// TwinCAT 3 PLC project TwinCAT_OpenFramework_Testing
// Title: TwinCAT Open Framework Testing
// Company: Oleksandr Tiutyk FOP
// Author: Oleksandr Tiutyk
// ProjectVersion: 1.0.13.0
// Description: Auumated testing engine implemenation
// ProgramVersion: 3.1.4026.28
// libraries:
//   Tc2_Utilities, * (Beckhoff Automation GmbH)
//   [TwinCAT Open Framework Core], * (Oleksandr Tiutyk FOP)
// project tree:
//   Assertions/ Assertions.TcPOU, AssertionContext.TcPOU
//   Assertions/TypedContexts/ BoolAssertionContext.TcPOU, SIntAssertionContext.TcPOU, IntAssertionContext.TcPOU, DIntAssertionContext.TcPOU, LIntAssertionContext.TcPOU, USIntAssertionContext.TcPOU, UIntAssertionContext.TcPOU, UDIntAssertionContext.TcPOU, ULIntAssertionContext.TcPOU, ByteAssertionContext.TcPOU, WordAssertionContext.TcPOU, DWordAssertionContext.TcPOU, LWordAssertionContext.TcPOU, RealAssertionContext.TcPOU, LongRealAssertionContext.TcPOU, StringAssertionContext.TcPOU, WideStringAssertionContext.TcPOU, TimeAssertionContext.TcPOU, LongTimeAssertionContext.TcPOU, DateAssertionContext.TcPOU, LongDateAssertionContext.TcPOU, DateTimeAssertionContext.TcPOU, LongDateTimeAssertionContext.TcPOU, TimeOfDayAssertionContext.TcPOU, LongTimeOfDayAssertionContext.TcPOU, PointerAssertionContext.TcPOU
//   Internal/ CurrentNamespace.TcPOU, NamespaceExtractor.TcPOU
//   Runner/ TEST_RUN_PHASE.TcDUT, TestRunner.TcPOU
//   TestElements/Groups/ TestGroup.TcPOU
//   TestElements/ IParentTestElement.TcIO, TEST_ELEMENT_STATE.TcDUT, ITestElement.TcIO, TestElement.TcPOU
//   TestElements/Tests/ TEST_CYCLE_RESULT.TcDUT, TEST_OUTCOME.TcDUT, ITestCase.TcIO, TestCase.TcPOU, SingleCycleTest.TcPOU, MultiCycleTest.TcPOU
//   Reporting/ ITestReporter.TcIO, AdsLogReporter.TcPOU, JUnitXmlReporter.TcPOU
//   / TestServices.TcPOU
//   Version/ Global_Version.TcGVL
// (motion and I/O tree: see PLC project twincat_openframework_core)
// real-time tasks:
//   TASK PlcTask: cycle T#10ms, priority 20, ADS port 350
//   TASK TestTask: cycle T#10ms, priority 1, ADS port 351
//   TASK RunnerTestTask: cycle T#10ms, priority 2, ADS port 354
//   TASK HowToTask: cycle T#10ms, priority 22, ADS port 353
// variable links:

// ---- Runner/TEST_RUN_PHASE.TcDUT
(*
SPDX-FileCopyrightText: © 2026 Oleksandr Tiutyk <trofimich@gmail.com>
SPDX-License-Identifier: MIT
License: https://opensource.org/license/mit
*)

(*!
<summary>Identifies the next root scheduling or reporting action.</summary>
*)

{attribute 'qualified_only'}
{attribute 'strict'}
{attribute 'to_string'}
TYPE TEST_RUN_PHASE :
(
	STARTING,
	RUNNING_ELEMENTS,
	REPORTING_TOTALS,
	COMPLETED
);
END_TYPE

// ---- TestElements/Tests/TEST_CYCLE_RESULT.TcDUT
(*
SPDX-FileCopyrightText: © 2026 Oleksandr Tiutyk <trofimich@gmail.com>
SPDX-License-Identifier: MIT
License: https://opensource.org/license/mit
*)

(*!
<summary>Indicates whether a test body needs more scheduling cycles or has finished on the current cycle.</summary>
<description>
BUSY (0) is the default uninitialized value and keeps the test running across subsequent cycles unless a failure
or deadline terminates the run. DONE (1) requests normal completion after the current cycle returns.
</description>
*)

{attribute 'qualified_only'}
{attribute 'strict'}
{attribute 'to_string'}
TYPE TEST_CYCLE_RESULT :
(
	BUSY := 0,
	DONE := 1
);
END_TYPE

// ---- TestElements/Tests/TEST_OUTCOME.TcDUT
(*
SPDX-FileCopyrightText: © 2026 Oleksandr Tiutyk <trofimich@gmail.com>
SPDX-License-Identifier: MIT
License: https://opensource.org/license/mit
*)

(*!
<summary>Defines the execution outcome of an individual test scenario.</summary>
<description>
Tracks whether a test has not yet run, is currently executing across cycles, passed all assertions, failed an
assertion or invariant, or was explicitly skipped.
</description>
*)

{attribute 'qualified_only'}
{attribute 'strict'}
{attribute 'to_string'}
TYPE TEST_OUTCOME :
(
	NOT_RUN := 0,
	RUNNING := 1,
	PASSED := 2,
	FAILED := 3,
	SKIPPED := 4
);
END_TYPE

// ---- TestElements/TEST_ELEMENT_STATE.TcDUT
(*
SPDX-FileCopyrightText: © 2026 Oleksandr Tiutyk <trofimich@gmail.com>
SPDX-License-Identifier: MIT
License: https://opensource.org/license/mit
*)

(*!
<summary>Identifies the execution lifecycle of a test element.</summary>
*)

{attribute 'qualified_only'}
{attribute 'strict'}
{attribute 'to_string'}
TYPE TEST_ELEMENT_STATE :
(
	READY,
	RUNNING,
	COMPLETED
);
END_TYPE

// ---- Version/Global_Version.TcGVL
{attribute 'TcGenerated'}
{attribute 'no-analysis'}
{attribute 'linkalways'}
// This function has been automatically generated from the project information.
VAR_GLOBAL CONSTANT
	{attribute 'const_non_replaced'}
	stLibVersion_TwinCAT_Open_Framework_Testing : ST_LibVersion := (iMajor := 1, iMinor := 0, iBuild := 13, iRevision := 0, nFlags := 0, sVersion := '1.0.13.0');
END_VAR

// ---- TestElements/IParentTestElement.TcIO
(*
SPDX-FileCopyrightText: © 2026 Oleksandr Tiutyk <trofimich@gmail.com>
SPDX-License-Identifier: MIT
License: https://opensource.org/license/mit
*)

(*!
<summary>Exposes borrowed direct children of a test element in fixed execution order.</summary>
<description>
ChildCount is stable throughout the element's lifetime; each direct child occupies one non-null slot.
GetChildByIndex borrows a child without resetting or executing it and transfers no allocation ownership.
Children and parent links obey ITestElement lifetime and lifecycle rules. Observations belong to the owning
task without reentry or cross-task synchronization. An empty composition has ChildCount zero and no valid index.
</description>
*)

INTERFACE IParentTestElement EXTENDS ITestElement

(*!
<summary>Reports the fixed number of direct children, including zero for an empty composition.</summary>
*)

{attribute 'monitoring' := 'call'}
PROPERTY FINAL ChildCount : TOF_Core.INT_LENGTH
GET
END_GET
END_PROPERTY

(*!
<summary>Borrows a direct child by its zero-based position in fixed execution order.</summary>
<description>
Available before the first Reset and after a failed Reset, provided the backing array and selected slot exist.
Missing storage or a null selected slot raises DataMemberNotSpecifiedException. Storage is checked first;
an index outside zero through ChildCount minus one raises ArgumentOutOfRangeException.
Does not mutate or execute the child, repeat whole-tree validation, or transfer ownership.
The child must remain alive while the interface is used; use only from the tree's owning task without reentry.
</description>
<param name="index">Zero-based direct-child position; an empty composition has no valid value.</param>
*)
METHOD GetChildByIndex : ITestElement
VAR_INPUT
	index : TOF_Core.INT_LENGTH;
END_VAR
END_METHOD

END_INTERFACE

// ---- Reporting/ITestReporter.TcIO
(*
SPDX-FileCopyrightText: © 2026 Oleksandr Tiutyk <trofimich@gmail.com>
SPDX-License-Identifier: MIT
License: https://opensource.org/license/mit
*)

(*!
<summary>Receives run boundaries and one terminal result per leaf test.</summary>
<description>
Callbacks execute synchronously in the owning runner task. Inputs are borrowed for the call only.
Do not retain them, reenter the tree, or share mutable reporter state between tasks. An exception aborts the
runner with ExitCode -1; output may be incomplete and the callback is not retried. Group paths are bounded
slash-separated display names. Groups do not emit synthetic test results or nested suite callbacks.
ReportTestCaseResult requires PASSED, FAILED or SKIPPED; other outcomes are invalid configuration.
Individual test names are bounded to 80 wide characters, matching INamed; group paths retain their 255-character bound.
</description>
*)

INTERFACE ITestReporter EXTENDS TOF_Core.IObject

(*!
<summary>Completes a run with aggregated leaf counts and nominal duration.</summary>
*)
METHOD ReportRunEnd
VAR_INPUT
	totalTests : TOF_Core.DINT_LENGTH;
	passedTests : TOF_Core.DINT_LENGTH;
	failedTests : TOF_Core.DINT_LENGTH;
	skippedTests : TOF_Core.DINT_LENGTH;
	duration : TIME;
END_VAR
END_METHOD

(*!
<summary>Begins a run with the number of configured leaf tests, including those that may be skipped.</summary>
<param name="testCount">The sum of the root TestCount values before executing any test.</param>
*)
METHOD ReportRunStart
VAR_INPUT
	testCount : TOF_Core.DINT_LENGTH;
END_VAR
END_METHOD

(*!
<summary>Receives one terminal leaf outcome and its first copied diagnostic.</summary>
<param name="testName">Individual name of at most 80 wide characters; longer input uses IEC truncation.</param>
*)
METHOD ReportTestCaseResult
VAR_INPUT
	groupPath : WSTRING(255);
	testName : WSTRING;
	outcome : TEST_OUTCOME;
	duration : TIME;
END_VAR
VAR_IN_OUT CONSTANT
	message : TOF_Core.ERROR_MESSAGE;
END_VAR
END_METHOD

END_INTERFACE

// ---- TestElements/ITestElement.TcIO
(*
SPDX-FileCopyrightText: © 2026 Oleksandr Tiutyk <trofimich@gmail.com>
SPDX-License-Identifier: MIT
License: https://opensource.org/license/mit
*)

(*!
<summary>Common cyclic execution contract for an individual test or a group of tests.</summary>
<description>
A live element occupies one slot of one tree. Its parent is assigned at construction and remains unchanged.
Its parent, descendants, reporter and tested resources remain alive and stable during a run.
All execution, configuration and observation of a tree belong to one cyclic task without reentry.
Separate tasks use disjoint trees, reporters and mutable tested resources; this interface provides no synchronization.
Execute advances at most one leaf body per call. A completed element ignores Execute until Reset.
Outcome counters describe leaf results. TestCount describes the configured leaf population of the subtree.
Custom implementations must preserve parent links and all lifecycle rules; callback exceptions abort the runner.
</description>
*)

INTERFACE ITestElement EXTENDS TOF_Core.INamed, TOF_Core.IExecutable

(*!
<summary>Reports nominal execution duration accumulated from calling task periods.</summary>
*)
{attribute 'monitoring' := 'call'}
PROPERTY Duration : TIME
GET
END_GET
END_PROPERTY

(*!
<summary>Counts failed leaf tests in this element.</summary>
*)
{attribute 'monitoring' := 'call'}
PROPERTY FailedCount : TOF_Core.DINT_LENGTH
GET
END_GET
END_PROPERTY

(*!
<summary>Builds the full display path from the root through this element.</summary>
<description>
Joins nonempty names with '/', including this element's name. A nameless root returns an empty path.
The result is a copied WSTRING bounded to 255 characters; overflow preserves the root prefix and ends with an ellipsis.
Reads the live Parent and Name properties without caching or changing the tree. All providers must remain alive
and stable during the call; use only in the owning task without reentry. Can be called before Reset.
A cyclic Parent chain raises StandardException to prevent an endless traversal. Provider exceptions propagate;
no element state or ownership is changed. Valid traversal uses fixed local strings without recursion or heap allocation.
</description>
*)
METHOD GetPath : WSTRING(255)
END_METHOD

(*!
<summary>Reports whether this element has completed.</summary>
*)
{attribute 'monitoring' := 'call'}
PROPERTY IsFinished : BOOL
GET
END_GET
END_PROPERTY

(*!
<summary>Reports whether this element has started and has not completed.</summary>
*)
{attribute 'monitoring' := 'call'}
PROPERTY IsRunning : BOOL
GET
END_GET
END_PROPERTY

(*!
<summary>Returns the group assigned at construction, or zero for a root.</summary>
<description>
Borrowed lifetime association. Reset and execution do not change it; the parent must remain alive.
Root registration with a runner does not bind Parent; a root must belong to one runner only.
</description>
*)
{attribute 'monitoring' := 'call'}
PROPERTY Parent : ITestElement
GET
END_GET
END_PROPERTY

(*!
<summary>Counts passed leaf tests in this element.</summary>
*)
{attribute 'monitoring' := 'call'}
PROPERTY PassedCount : TOF_Core.DINT_LENGTH
GET
END_GET
END_PROPERTY

(*!
<summary>Reports nominal scheduled duration, not CPU execution time.</summary>
*)
{attribute 'monitoring' := 'call'}
PROPERTY FINAL Reporter : ITestReporter
GET
END_GET
END_PROPERTY

(*!
<summary>Prepares a fresh run and borrows the reporter.</summary>
<description>
Call before first execution, after completion, or after an aborted run once resources are safe.
This is not cancellation: it does not execute test teardown. The reporter may be zero to suppress reporting.
Group reset recursively resets descendants. External callback exceptions propagate; partial reset is possible.
</description>
*)
METHOD Reset
VAR_INPUT
	reporter : ITestReporter;
END_VAR
END_METHOD

(*!
<summary>Counts skipped leaf tests in this element.</summary>
*)
{attribute 'monitoring' := 'call'}
PROPERTY SkippedCount : TOF_Core.DINT_LENGTH
GET
END_GET
END_PROPERTY

(*!
<summary>Reports nominal scheduled duration, not CPU execution time.</summary>
*)
{attribute 'monitoring' := 'call'}
PROPERTY FINAL State : TEST_ELEMENT_STATE
GET
END_GET
END_PROPERTY

(*!
<summary>Counts the configured leaf tests in this subtree.</summary>
<description>
A leaf counts as one regardless of its outcome. Groups sum their children; an empty group counts as zero.
Read from the owning task after the tree has been constructed. The caller supplies a valid, stable subtree
whose total fits in UDINT. Reading does not run or reset tests, and the value is stable across runs.
Provider exceptions propagate.
</description>
*)
{attribute 'monitoring' := 'call'}
PROPERTY TestCount : TOF_Core.DINT_LENGTH
GET
END_GET
END_PROPERTY

END_INTERFACE

// ---- TestElements/Tests/ITestCase.TcIO
(*
SPDX-FileCopyrightText: © 2026 Oleksandr Tiutyk <trofimich@gmail.com>
SPDX-License-Identifier: MIT
License: https://opensource.org/license/mit
*)

(*!
<summary>Receives assertion failures for one individual test.</summary>
<description>
Groups use ITestElement and do not receive leaf assertions. A failure is copied only while the case is running.
</description>
*)

INTERFACE ITestCase EXTENDS ITestElement

(*!
<summary>Copies the first failure of the running case; later diagnostics do not replace it.</summary>
*)
METHOD RecordFailure
VAR_IN_OUT CONSTANT
	message : TOF_Core.ERROR_MESSAGE;
END_VAR
END_METHOD

END_INTERFACE

// ---- Assertions/Assertions.TcPOU
(*
SPDX-FileCopyrightText: © 2026 Oleksandr Tiutyk <trofimich@gmail.com>
SPDX-License-Identifier: MIT
License: https://opensource.org/license/mit
*)

(*!
<summary>Provides fluent test assertion entry points on values, variables, and objects.</summary>
<description>
TestCase owns and binds this instance before its first callback.
Typed That methods copy actual values into independent persistent contexts; generic That borrows a live variable.
Contexts do not call one another; shared services only report failures and implement floating value policy.
Finish one immediate chain before starting another, regardless of operand type. Do not retain a returned
context or use this provider across tasks or reentrantly. Every entry verifies that its owning case is running.
An optional copied message prefixes every assertion failure in the chain and is replaced on the next entry.
Typed contexts apply ordinary IEC input conversions; select the entry matching the intended operand type.
Do not copy this provider by value: its contexts retain borrowed links to the owning test case and actual storage.
</description>
*)

{attribute 'no_explicit_call' := 'do not call this function block directly'}
FUNCTION_BLOCK Assertions EXTENDS TOF_Core.Object
VAR_STAT
	{attribute 'hide'} 
	_ClassName : STRING := __POUNAME();	
END_VAR
VAR	
	_AssertionContext : AssertionContext;
	
	_BoolContext : BoolAssertionContext;
	_SIntContext : SIntAssertionContext;
	_IntContext : IntAssertionContext;
	_DIntContext : DIntAssertionContext;
	_LIntContext : LIntAssertionContext;
	_USIntContext : USIntAssertionContext;
	_UIntContext : UIntAssertionContext;
	_UDIntContext : UDIntAssertionContext;
	_ULIntContext : ULIntAssertionContext;
	_ByteContext : ByteAssertionContext;
	_WordContext : WordAssertionContext;
	_DWordContext : DWordAssertionContext;
	_LWordContext : LWordAssertionContext;
	_RealContext : RealAssertionContext;
	_LongRealContext : LongRealAssertionContext;
	_StringContext : StringAssertionContext;
	_WideStringContext : WideStringAssertionContext;
	_TimeContext : TimeAssertionContext;
	_LongTimeContext : LongTimeAssertionContext;
	_DateContext : DateAssertionContext;
	_LongDateContext : LongDateAssertionContext;
	_DateTimeContext : DateTimeAssertionContext;
	_LongDateTimeContext : LongDateTimeAssertionContext;
	_TimeOfDayContext : TimeOfDayAssertionContext;
	_LongTimeOfDayContext : LongTimeOfDayAssertionContext;
	_PointerContext : PointerAssertionContext;
	
	_TestCase : ITestCase;
END_VAR

//! <summary>Borrows the owning test case for assertion failure reporting throughout the run.</summary>
METHOD INTERNAL FINAL Bind
VAR_INPUT
	testCase : ITestCase;
END_VAR
_TestCase := testCase;
END_METHOD

//! <summary>Provides assertion-provider metadata.</summary>
{attribute 'monitoring' := 'call'}
PROPERTY ClassName : REFERENCE TO STRING
GET
ClassName REF= _ClassName;
END_GET
END_PROPERTY

(*!
<summary>Returns the namespace name of this assertion provider.</summary>
*)
{attribute 'monitoring' := 'call'}
PROPERTY NamespaceName : REFERENCE TO STRING
GET
NamespaceName REF= CurrentNamespace.Name;
END_GET
END_PROPERTY

(*!
<summary>Rejects assertion entry outside a running owning case before context mutation.</summary>
<description>
Raises DataMemberNotSpecifiedException when no running test case is bound.
</description>
*)
METHOD PRIVATE requireRunningCase
IF _TestCase = 0 OR_ELSE NOT _TestCase.IsRunning THEN
	TOF_Core.Exceptions.ThrowDataMemberNotSpecified(
		sourceNamespaceName := NamespaceName,
		sourceClassName := ClassName,
		sourcePOUName := __POUNAME(),
		sourcePosition := __POSITION(),
		dataMemberName := '_TestCase'
	);
END_IF
END_METHOD

(*!
<summary>Reports the byte size of this concrete instance.</summary>
<description>
Uses XSIZEOF on the instance. Does not include separately allocated payloads or prove that an arbitrary
address is valid.
</description>
*)
{attribute 'monitoring' := 'call'}
PROPERTY SelfSize : ULINT
GET
SelfSize := XSIZEOF(THIS^);
END_GET
END_PROPERTY

(*!
<summary>Begins a fluent assertion chain on the provided actual value.</summary>
<description>
Borrows actual storage for this expression; actual must be a variable. Use typed entry points for literals
and expression results. Starting another chain replaces that entry's operand and message.
Calling That without a running owning case raises DataMemberNotSpecifiedException.
Equality follows GENERIC_VALUE byte/value semantics; FB operands do not invoke Object.Equals.
For object equality, use ThatBool on the Boolean result of its explicit Equals call.
</description>
<param name="actual">Live variable borrowed through the immediate chain.</param>
<param name="message">Optional copied prefix for every failure in this chain; default empty.</param>
*)
METHOD That : REFERENCE TO AssertionContext
VAR_INPUT
	actual : ANY;
	message : WSTRING(255) := "";
END_VAR
requireRunningCase();

_AssertionContext.Prepare(actual := actual, testCase := _TestCase, message := message);

That REF= _AssertionContext;
END_METHOD

(*!
<summary>Begins a fluent chain on a copied BOOL value.</summary>
<description>
Accepts literals, variables and expression results through a concrete IEC input type.
Requires a running owning case; otherwise raises DataMemberNotSpecifiedException.
Finish this chain before starting another. The message applies to every assertion in the chain.
</description>
<param name="actual">Value copied after ordinary IEC conversion to BOOL.</param>
<param name="message">Optional copied diagnostic prefix; default empty replaces the previous prefix.</param>
*)
METHOD ThatBool : REFERENCE TO BoolAssertionContext
VAR_INPUT
	actual : BOOL;
	message : WSTRING(255) := "";
END_VAR
requireRunningCase();

_BoolContext.Prepare(actual := actual, testCase := _TestCase, message := message);

ThatBool REF= _BoolContext;
END_METHOD

(*!
<summary>Begins a fluent chain on a copied BYTE value.</summary>
<description>
Accepts literals, variables and expression results through a concrete IEC input type.
Requires a running owning case; otherwise raises DataMemberNotSpecifiedException.
Finish this chain before starting another. The message applies to every assertion in the chain.
</description>
<param name="actual">Value copied after ordinary IEC conversion to BYTE.</param>
<param name="message">Optional copied diagnostic prefix; default empty replaces the previous prefix.</param>
*)
METHOD ThatByte : REFERENCE TO ByteAssertionContext
VAR_INPUT
	actual : BYTE;
	message : WSTRING(255) := "";
END_VAR
requireRunningCase();

_ByteContext.Prepare(actual := actual, testCase := _TestCase, message := message);

ThatByte REF= _ByteContext;
END_METHOD

(*!
<summary>Begins a fluent chain on a copied DATE value.</summary>
<description>
Accepts literals, variables and expression results through a concrete IEC input type.
Requires a running owning case; otherwise raises DataMemberNotSpecifiedException.
Finish this chain before starting another. The message applies to every assertion in the chain.
</description>
<param name="actual">Value copied after ordinary IEC conversion to DATE.</param>
<param name="message">Optional copied diagnostic prefix; default empty replaces the previous prefix.</param>
*)
METHOD ThatDate : REFERENCE TO DateAssertionContext
VAR_INPUT
	actual : DATE;
	message : WSTRING(255) := "";
END_VAR
requireRunningCase();

_DateContext.Prepare(actual := actual, testCase := _TestCase, message := message);

ThatDate REF= _DateContext;
END_METHOD

(*!
<summary>Begins a fluent chain on a copied DATE_AND_TIME value.</summary>
<description>
Accepts literals, variables and expression results through a concrete IEC input type.
Requires a running owning case; otherwise raises DataMemberNotSpecifiedException.
Finish this chain before starting another. The message applies to every assertion in the chain.
</description>
<param name="actual">Value copied after ordinary IEC conversion to DATE_AND_TIME.</param>
<param name="message">Optional copied diagnostic prefix; default empty replaces the previous prefix.</param>
*)
METHOD ThatDateTime : REFERENCE TO DateTimeAssertionContext
VAR_INPUT
	actual : DATE_AND_TIME;
	message : WSTRING(255) := "";
END_VAR
requireRunningCase();

_DateTimeContext.Prepare(actual := actual, testCase := _TestCase, message := message);

ThatDateTime REF= _DateTimeContext;
END_METHOD

(*!
<summary>Begins a fluent chain on a copied DINT value.</summary>
<description>
Accepts literals, variables and expression results through a concrete IEC input type.
Requires a running owning case; otherwise raises DataMemberNotSpecifiedException.
Finish this chain before starting another. The message applies to every assertion in the chain.
</description>
<param name="actual">Value copied after ordinary IEC conversion to DINT.</param>
<param name="message">Optional copied diagnostic prefix; default empty replaces the previous prefix.</param>
*)
METHOD ThatDInt : REFERENCE TO DIntAssertionContext
VAR_INPUT
	actual : DINT;
	message : WSTRING(255) := "";
END_VAR
requireRunningCase();

_DIntContext.Prepare(actual := actual, testCase := _TestCase, message := message);

ThatDInt REF= _DIntContext;
END_METHOD

(*!
<summary>Begins a fluent chain on a copied DWORD value.</summary>
<description>
Accepts literals, variables and expression results through a concrete IEC input type.
Requires a running owning case; otherwise raises DataMemberNotSpecifiedException.
Finish this chain before starting another. The message applies to every assertion in the chain.
</description>
<param name="actual">Value copied after ordinary IEC conversion to DWORD.</param>
<param name="message">Optional copied diagnostic prefix; default empty replaces the previous prefix.</param>
*)
METHOD ThatDWord : REFERENCE TO DWordAssertionContext
VAR_INPUT
	actual : DWORD;
	message : WSTRING(255) := "";
END_VAR
requireRunningCase();

_DWordContext.Prepare(actual := actual, testCase := _TestCase, message := message);

ThatDWord REF= _DWordContext;
END_METHOD

(*!
<summary>Begins a fluent chain on a copied INT value.</summary>
<description>
Accepts literals, variables and expression results through a concrete IEC input type.
Requires a running owning case; otherwise raises DataMemberNotSpecifiedException.
Finish this chain before starting another. The message applies to every assertion in the chain.
</description>
<param name="actual">Value copied after ordinary IEC conversion to INT.</param>
<param name="message">Optional copied diagnostic prefix; default empty replaces the previous prefix.</param>
*)
METHOD ThatInt : REFERENCE TO IntAssertionContext
VAR_INPUT
	actual : INT;
	message : WSTRING(255) := "";
END_VAR
requireRunningCase();

_IntContext.Prepare(actual := actual, testCase := _TestCase, message := message);

ThatInt REF= _IntContext;
END_METHOD

(*!
<summary>Begins a fluent chain on a copied LINT value.</summary>
<description>
Accepts literals, variables and expression results through a concrete IEC input type.
Requires a running owning case; otherwise raises DataMemberNotSpecifiedException.
Finish this chain before starting another. The message applies to every assertion in the chain.
</description>
<param name="actual">Value copied after ordinary IEC conversion to LINT.</param>
<param name="message">Optional copied diagnostic prefix; default empty replaces the previous prefix.</param>
*)
METHOD ThatLInt : REFERENCE TO LIntAssertionContext
VAR_INPUT
	actual : LINT;
	message : WSTRING(255) := "";
END_VAR
requireRunningCase();

_LIntContext.Prepare(actual := actual, testCase := _TestCase, message := message);

ThatLInt REF= _LIntContext;
END_METHOD

(*!
<summary>Begins a fluent chain on a copied LDATE value.</summary>
<description>
Accepts literals, variables and expression results through a concrete IEC input type.
Requires a running owning case; otherwise raises DataMemberNotSpecifiedException.
Finish this chain before starting another. The message applies to every assertion in the chain.
</description>
<param name="actual">Value copied after ordinary IEC conversion to LDATE.</param>
<param name="message">Optional copied diagnostic prefix; default empty replaces the previous prefix.</param>
*)
METHOD ThatLongDate : REFERENCE TO LongDateAssertionContext
VAR_INPUT
	actual : LDATE;
	message : WSTRING(255) := "";
END_VAR
requireRunningCase();

_LongDateContext.Prepare(actual := actual, testCase := _TestCase, message := message);

ThatLongDate REF= _LongDateContext;
END_METHOD

(*!
<summary>Begins a fluent chain on a copied LDATE_AND_TIME value.</summary>
<description>
Accepts literals, variables and expression results through a concrete IEC input type.
Requires a running owning case; otherwise raises DataMemberNotSpecifiedException.
Finish this chain before starting another. The message applies to every assertion in the chain.
</description>
<param name="actual">Value copied after ordinary IEC conversion to LDATE_AND_TIME.</param>
<param name="message">Optional copied diagnostic prefix; default empty replaces the previous prefix.</param>
*)
METHOD ThatLongDateTime : REFERENCE TO LongDateTimeAssertionContext
VAR_INPUT
	actual : LDATE_AND_TIME;
	message : WSTRING(255) := "";
END_VAR
requireRunningCase();

_LongDateTimeContext.Prepare(actual := actual, testCase := _TestCase, message := message);

ThatLongDateTime REF= _LongDateTimeContext;
END_METHOD

(*!
<summary>Begins a fluent chain on a copied LREAL value.</summary>
<description>
Accepts literals, variables and expression results through a concrete IEC input type.
Requires a running owning case; otherwise raises DataMemberNotSpecifiedException.
Finish this chain before starting another. The message applies to every assertion in the chain.
</description>
<param name="actual">Value copied after ordinary IEC conversion to LREAL.</param>
<param name="message">Optional copied diagnostic prefix; default empty replaces the previous prefix.</param>
*)
METHOD ThatLongReal : REFERENCE TO LongRealAssertionContext
VAR_INPUT
	actual : LREAL;
	message : WSTRING(255) := "";
END_VAR
requireRunningCase();

_LongRealContext.Prepare(actual := actual, testCase := _TestCase, message := message);

ThatLongReal REF= _LongRealContext;
END_METHOD

(*!
<summary>Begins a fluent chain on a copied LTIME value.</summary>
<description>
Accepts literals, variables and expression results through a concrete IEC input type.
Requires a running owning case; otherwise raises DataMemberNotSpecifiedException.
Finish this chain before starting another. The message applies to every assertion in the chain.
</description>
<param name="actual">Value copied after ordinary IEC conversion to LTIME.</param>
<param name="message">Optional copied diagnostic prefix; default empty replaces the previous prefix.</param>
*)
METHOD ThatLongTime : REFERENCE TO LongTimeAssertionContext
VAR_INPUT
	actual : LTIME;
	message : WSTRING(255) := "";
END_VAR
requireRunningCase();

_LongTimeContext.Prepare(actual := actual, testCase := _TestCase, message := message);

ThatLongTime REF= _LongTimeContext;
END_METHOD

(*!
<summary>Begins a fluent chain on a copied LTIME_OF_DAY value.</summary>
<description>
Accepts literals, variables and expression results through a concrete IEC input type.
Requires a running owning case; otherwise raises DataMemberNotSpecifiedException.
Finish this chain before starting another. The message applies to every assertion in the chain.
</description>
<param name="actual">Value copied after ordinary IEC conversion to LTIME_OF_DAY.</param>
<param name="message">Optional copied diagnostic prefix; default empty replaces the previous prefix.</param>
*)
METHOD ThatLongTimeOfDay : REFERENCE TO LongTimeOfDayAssertionContext
VAR_INPUT
	actual : LTIME_OF_DAY;
	message : WSTRING(255) := "";
END_VAR
requireRunningCase();

_LongTimeOfDayContext.Prepare(actual := actual, testCase := _TestCase, message := message);

ThatLongTimeOfDay REF= _LongTimeOfDayContext;
END_METHOD

(*!
<summary>Begins a fluent chain on a copied LWORD value.</summary>
<description>
Accepts literals, variables and expression results through a concrete IEC input type.
Requires a running owning case; otherwise raises DataMemberNotSpecifiedException.
Finish this chain before starting another. The message applies to every assertion in the chain.
</description>
<param name="actual">Value copied after ordinary IEC conversion to LWORD.</param>
<param name="message">Optional copied diagnostic prefix; default empty replaces the previous prefix.</param>
*)
METHOD ThatLWord : REFERENCE TO LWordAssertionContext
VAR_INPUT
	actual : LWORD;
	message : WSTRING(255) := "";
END_VAR
requireRunningCase();

_LWordContext.Prepare(actual := actual, testCase := _TestCase, message := message);

ThatLWord REF= _LWordContext;
END_METHOD

(*!
<summary>Begins a fluent chain on a copied PVOID value.</summary>
<description>
Accepts literals, variables and expression results through a concrete IEC input type.
Requires a running owning case; otherwise raises DataMemberNotSpecifiedException.
Finish this chain before starting another. The message applies to every assertion in the chain.
</description>
<param name="actual">Value copied after ordinary IEC conversion to PVOID.</param>
<param name="message">Optional copied diagnostic prefix; default empty replaces the previous prefix.</param>
*)
METHOD ThatPointer : REFERENCE TO PointerAssertionContext
VAR_INPUT
	actual : PVOID;
	message : WSTRING(255) := "";
END_VAR
requireRunningCase();

_PointerContext.Prepare(actual := actual, testCase := _TestCase, message := message);

ThatPointer REF= _PointerContext;
END_METHOD

(*!
<summary>Begins a fluent chain on a copied REAL value.</summary>
<description>
Accepts literals, variables and expression results through a concrete IEC input type.
Requires a running owning case; otherwise raises DataMemberNotSpecifiedException.
Finish this chain before starting another. The message applies to every assertion in the chain.
</description>
<param name="actual">Value copied after ordinary IEC conversion to REAL.</param>
<param name="message">Optional copied diagnostic prefix; default empty replaces the previous prefix.</param>
*)
METHOD ThatReal : REFERENCE TO RealAssertionContext
VAR_INPUT
	actual : REAL;
	message : WSTRING(255) := "";
END_VAR
requireRunningCase();

_RealContext.Prepare(actual := actual, testCase := _TestCase, message := message);

ThatReal REF= _RealContext;
END_METHOD

(*!
<summary>Begins a fluent chain on a copied SINT value.</summary>
<description>
Accepts literals, variables and expression results through a concrete IEC input type.
Requires a running owning case; otherwise raises DataMemberNotSpecifiedException.
Finish this chain before starting another. The message applies to every assertion in the chain.
</description>
<param name="actual">Value copied after ordinary IEC conversion to SINT.</param>
<param name="message">Optional copied diagnostic prefix; default empty replaces the previous prefix.</param>
*)
METHOD ThatSInt : REFERENCE TO SIntAssertionContext
VAR_INPUT
	actual : SINT;
	message : WSTRING(255) := "";
END_VAR
requireRunningCase();

_SIntContext.Prepare(actual := actual, testCase := _TestCase, message := message);

ThatSInt REF= _SIntContext;
END_METHOD

(*!
<summary>Begins a fluent chain on a copied STRING(255) value.</summary>
<description>
Accepts literals, variables and expression results through a concrete IEC input type.
Requires a running owning case; otherwise raises DataMemberNotSpecifiedException.
Inputs are bounded to 255 characters. Finish this chain before starting another.
The message applies to every assertion in the chain.
</description>
<param name="actual">Value copied after ordinary IEC conversion to STRING(255).</param>
<param name="message">Optional copied diagnostic prefix; default empty replaces the previous prefix.</param>
*)
METHOD ThatString : REFERENCE TO StringAssertionContext
VAR_INPUT
	actual : STRING(255);
	message : WSTRING(255) := "";
END_VAR
requireRunningCase();

_StringContext.Prepare(actual := actual, testCase := _TestCase, message := message);

ThatString REF= _StringContext;
END_METHOD

(*!
<summary>Begins a fluent chain on a copied TIME value.</summary>
<description>
Accepts literals, variables and expression results through a concrete IEC input type.
Requires a running owning case; otherwise raises DataMemberNotSpecifiedException.
Finish this chain before starting another. The message applies to every assertion in the chain.
</description>
<param name="actual">Value copied after ordinary IEC conversion to TIME.</param>
<param name="message">Optional copied diagnostic prefix; default empty replaces the previous prefix.</param>
*)
METHOD ThatTime : REFERENCE TO TimeAssertionContext
VAR_INPUT
	actual : TIME;
	message : WSTRING(255) := "";
END_VAR
requireRunningCase();

_TimeContext.Prepare(actual := actual, testCase := _TestCase, message := message);

ThatTime REF= _TimeContext;
END_METHOD

(*!
<summary>Begins a fluent chain on a copied TIME_OF_DAY value.</summary>
<description>
Accepts literals, variables and expression results through a concrete IEC input type.
Requires a running owning case; otherwise raises DataMemberNotSpecifiedException.
Finish this chain before starting another. The message applies to every assertion in the chain.
</description>
<param name="actual">Value copied after ordinary IEC conversion to TIME_OF_DAY.</param>
<param name="message">Optional copied diagnostic prefix; default empty replaces the previous prefix.</param>
*)
METHOD ThatTimeOfDay : REFERENCE TO TimeOfDayAssertionContext
VAR_INPUT
	actual : TIME_OF_DAY;
	message : WSTRING(255) := "";
END_VAR
requireRunningCase();

_TimeOfDayContext.Prepare(actual := actual, testCase := _TestCase, message := message);

ThatTimeOfDay REF= _TimeOfDayContext;
END_METHOD

(*!
<summary>Begins a fluent chain on a copied UDINT value.</summary>
<description>
Accepts literals, variables and expression results through a concrete IEC input type.
Requires a running owning case; otherwise raises DataMemberNotSpecifiedException.
Finish this chain before starting another. The message applies to every assertion in the chain.
</description>
<param name="actual">Value copied after ordinary IEC conversion to UDINT.</param>
<param name="message">Optional copied diagnostic prefix; default empty replaces the previous prefix.</param>
*)
METHOD ThatUDInt : REFERENCE TO UDIntAssertionContext
VAR_INPUT
	actual : UDINT;
	message : WSTRING(255) := "";
END_VAR
requireRunningCase();

_UDIntContext.Prepare(actual := actual, testCase := _TestCase, message := message);

ThatUDInt REF= _UDIntContext;
END_METHOD

(*!
<summary>Begins a fluent chain on a copied UINT value.</summary>
<description>
Accepts literals, variables and expression results through a concrete IEC input type.
Requires a running owning case; otherwise raises DataMemberNotSpecifiedException.
Finish this chain before starting another. The message applies to every assertion in the chain.
</description>
<param name="actual">Value copied after ordinary IEC conversion to UINT.</param>
<param name="message">Optional copied diagnostic prefix; default empty replaces the previous prefix.</param>
*)
METHOD ThatUInt : REFERENCE TO UIntAssertionContext
VAR_INPUT
	actual : UINT;
	message : WSTRING(255) := "";
END_VAR
requireRunningCase();

_UIntContext.Prepare(actual := actual, testCase := _TestCase, message := message);

ThatUInt REF= _UIntContext;
END_METHOD

(*!
<summary>Begins a fluent chain on a copied ULINT value.</summary>
<description>
Accepts literals, variables and expression results through a concrete IEC input type.
Requires a running owning case; otherwise raises DataMemberNotSpecifiedException.
Finish this chain before starting another. The message applies to every assertion in the chain.
</description>
<param name="actual">Value copied after ordinary IEC conversion to ULINT.</param>
<param name="message">Optional copied diagnostic prefix; default empty replaces the previous prefix.</param>
*)
METHOD ThatULInt : REFERENCE TO ULIntAssertionContext
VAR_INPUT
	actual : ULINT;
	message : WSTRING(255) := "";
END_VAR
requireRunningCase();

_ULIntContext.Prepare(actual := actual, testCase := _TestCase, message := message);

ThatULInt REF= _ULIntContext;
END_METHOD

(*!
<summary>Begins a fluent chain on a copied USINT value.</summary>
<description>
Accepts literals, variables and expression results through a concrete IEC input type.
Requires a running owning case; otherwise raises DataMemberNotSpecifiedException.
Finish this chain before starting another. The message applies to every assertion in the chain.
</description>
<param name="actual">Value copied after ordinary IEC conversion to USINT.</param>
<param name="message">Optional copied diagnostic prefix; default empty replaces the previous prefix.</param>
*)
METHOD ThatUSInt : REFERENCE TO USIntAssertionContext
VAR_INPUT
	actual : USINT;
	message : WSTRING(255) := "";
END_VAR
requireRunningCase();

_USIntContext.Prepare(actual := actual, testCase := _TestCase, message := message);

ThatUSInt REF= _USIntContext;
END_METHOD

(*!
<summary>Begins a fluent chain on a copied WSTRING(255) value.</summary>
<description>
Accepts literals, variables and expression results through a concrete IEC input type.
Requires a running owning case; otherwise raises DataMemberNotSpecifiedException.
Inputs are bounded to 255 characters. Finish this chain before starting another.
The message applies to every assertion in the chain.
</description>
<param name="actual">Value copied after ordinary IEC conversion to WSTRING(255).</param>
<param name="message">Optional copied diagnostic prefix; default empty replaces the previous prefix.</param>
*)
METHOD ThatWideString : REFERENCE TO WideStringAssertionContext
VAR_INPUT
	actual : WSTRING(255);
	message : WSTRING(255) := "";
END_VAR
requireRunningCase();

_WideStringContext.Prepare(actual := actual, testCase := _TestCase, message := message);

ThatWideString REF= _WideStringContext;
END_METHOD

(*!
<summary>Begins a fluent chain on a copied WORD value.</summary>
<description>
Accepts literals, variables and expression results through a concrete IEC input type.
Requires a running owning case; otherwise raises DataMemberNotSpecifiedException.
Finish this chain before starting another. The message applies to every assertion in the chain.
</description>
<param name="actual">Value copied after ordinary IEC conversion to WORD.</param>
<param name="message">Optional copied diagnostic prefix; default empty replaces the previous prefix.</param>
*)
METHOD ThatWord : REFERENCE TO WordAssertionContext
VAR_INPUT
	actual : WORD;
	message : WSTRING(255) := "";
END_VAR
requireRunningCase();

_WordContext.Prepare(actual := actual, testCase := _TestCase, message := message);

ThatWord REF= _WordContext;
END_METHOD

END_FUNCTION_BLOCK

// ---- Assertions/AssertionContext.TcPOU
(*
SPDX-FileCopyrightText: © 2026 Oleksandr Tiutyk <trofimich@gmail.com>
SPDX-License-Identifier: MIT
License: https://opensource.org/license/mit
*)

(*!
<summary>Provides a fluent assertion builder for polymorphic value and reference assertions.</summary>
<description>
Borrows actual storage for one immediate assertion chain on one task. Use inside a running test callback.
ANY operands must be variables; use the typed That methods for literals, expressions and property results.
The copied message prefixes every failure in this chain until Prepare starts another chain.
The test case retains the first failure without interrupting the callback.
Equality uses GENERIC_VALUE.Equals: integer widths/signedness compare by value; floating values use canonical
equality; unlike type categories remain distinct. USER_DEFINED/FB values compare stored bytes, including
padding and aliases, not Object.Equals. Use ThatBool on an explicit Equals result for object equality.
Pointer equality compares pointer values, not pointed-to contents. Public generic comparisons are exact;
only the independent typed REAL/LREAL contexts expose absolute tolerance arguments.
Unsupported conversions may raise framework exceptions. No cross-task use or same-instance reentry is supported.
</description>
*)

{attribute 'no_explicit_call' := 'do not call this function block directly'}
FUNCTION_BLOCK AssertionContext EXTENDS TOF_Core.Object
VAR_STAT
	{attribute 'hide'} 
	_ClassName : STRING := __POUNAME();
END_VAR
VAR
	_TestCase : ITestCase;
	_Actual : TOF_Core.GENERIC_VALUE;	
	_Message : WSTRING(255);
END_VAR

//! <summary>Provides assertion-context metadata.</summary>
{attribute 'monitoring' := 'call'}
PROPERTY ClassName : REFERENCE TO STRING
GET
ClassName REF= _ClassName;
END_GET
END_PROPERTY

(*!
<summary>Reports to the bound test case with the current chain message.</summary>
<description>
A missing receiver raises DataMemberNotSpecifiedException. Shared reporting retains no context state;
receiver exceptions propagate to the enclosing test callback handler.
</description>
<param name="defaultMessage">Diagnostic borrowed only during reporting.</param>
*)
METHOD PRIVATE fail
VAR_IN_OUT CONSTANT
	defaultMessage : TOF_Core.ERROR_MESSAGE;
END_VAR
TestServices.ReportAssertionFailure(
	testCase := _TestCase,
	message := _Message,
	sourceClassName := ClassName,
	defaultMessage := defaultMessage
);
END_METHOD

(*!
<summary>Asserts that the actual value is a boolean equal to FALSE.</summary>
<description>
A non-Boolean operand or TRUE records failure; the chain message remains available.
</description>
*)
METHOD FINAL IsFalse : REFERENCE TO AssertionContext
VAR
	diagnostic : TOF_Core.ERROR_MESSAGE;
END_VAR
IF _Actual.TypeClass <> TOF_Core.GENERIC_TYPE_CLASS.BOOLEAN OR_ELSE _Actual.AsBool() THEN
	diagnostic := TOF_Core.WideStrings.Concat255(
		"Expected: FALSE, but was: ",
		_Actual.AsWString255()
	);
	fail(defaultMessage := diagnostic);
END_IF

IsFalse REF= THIS^;
END_METHOD

(*!
<summary>Asserts that the actual value is strictly greater than the expected variable.</summary>
<description>
Uses Core ordering without tolerance. Comparison exceptions record an assertion failure.
The chain message remains available to subsequent assertions.
</description>
<param name="expected">Live variable to compare; ANY does not accept literals or expression results.</param>
*)
METHOD FINAL IsGreaterThan : REFERENCE TO AssertionContext
VAR_INPUT
	expected : ANY;
END_VAR
VAR
	diagnostic : TOF_Core.ERROR_MESSAGE;
	expectedGeneric : TOF_Core.GENERIC_VALUE;
	comparison : TOF_Core.COMPARISON_RESULT;
	isOrdered : BOOL;
END_VAR
expectedGeneric := TOF_Core.GenericValueFactory.FromAny(
	value := expected,
	isObject := FALSE,
	memoryManagementBehavior := TOF_Core.GENERIC_MEMORY_MANAGEMENT_BEHAVIOR.STORE_ORIGINAL_REFERENCE_AND_NOT_OWNS_MEMORY
);

__TRY
	comparison := _Actual.CompareTo(otherValue := expectedGeneric);
	isOrdered := (comparison = TOF_Core.COMPARISON_RESULT.FIRST_GREATER_THAN_SECOND);
__CATCH
	isOrdered := FALSE;
__ENDTRY

IF NOT isOrdered THEN
	diagnostic := TOF_Core.WideStrings.Concat255(
		"Expected value > ",
		expectedGeneric.AsWString255(),
		", but was: ",
		_Actual.AsWString255()
	);
	fail(defaultMessage := diagnostic);
END_IF

IsGreaterThan REF= THIS^;
END_METHOD

(*!
<summary>Asserts that the actual value meets the inclusive lower boundary.</summary>
<description>
Uses Core ordering without tolerance. Comparison exceptions record an assertion failure.
The chain message remains available to subsequent assertions.
</description>
<param name="expected">Live variable to compare; ANY does not accept literals or expression results.</param>
*)
METHOD FINAL IsGreaterThanOrEquals : REFERENCE TO AssertionContext
VAR_INPUT
	expected : ANY;
END_VAR
VAR
	diagnostic : TOF_Core.ERROR_MESSAGE;
	expectedGeneric : TOF_Core.GENERIC_VALUE;
	comparison : TOF_Core.COMPARISON_RESULT;
	isOrdered : BOOL;
END_VAR
expectedGeneric := TOF_Core.GenericValueFactory.FromAny(
	value := expected,
	isObject := FALSE,
	memoryManagementBehavior := TOF_Core.GENERIC_MEMORY_MANAGEMENT_BEHAVIOR.STORE_ORIGINAL_REFERENCE_AND_NOT_OWNS_MEMORY
);

__TRY
	comparison := _Actual.CompareTo(otherValue := expectedGeneric);
	isOrdered := (comparison = TOF_Core.COMPARISON_RESULT.FIRST_GREATER_THAN_SECOND)
		OR_ELSE (comparison = TOF_Core.COMPARISON_RESULT.FIRST_EQUAL_TO_SECOND);
__CATCH
	isOrdered := FALSE;
__ENDTRY

IF NOT isOrdered THEN
	diagnostic := TOF_Core.WideStrings.Concat255(
		"Expected value >= ",
		expectedGeneric.AsWString255(),
		", but was: ",
		_Actual.AsWString255()
	);
	fail(defaultMessage := diagnostic);
END_IF

IsGreaterThanOrEquals REF= THIS^;
END_METHOD

(*!
<summary>Asserts that the actual value is strictly less than the expected variable.</summary>
<description>
Uses Core ordering without tolerance. Comparison exceptions record an assertion failure.
The chain message remains available to subsequent assertions.
</description>
<param name="expected">Live variable to compare; ANY does not accept literals or expression results.</param>
*)
METHOD FINAL IsLessThan : REFERENCE TO AssertionContext
VAR_INPUT
	expected : ANY;
END_VAR
VAR
	diagnostic : TOF_Core.ERROR_MESSAGE;
	expectedGeneric : TOF_Core.GENERIC_VALUE;
	comparison : TOF_Core.COMPARISON_RESULT;
	isOrdered : BOOL;
END_VAR
expectedGeneric := TOF_Core.GenericValueFactory.FromAny(
	value := expected,
	isObject := FALSE,
	memoryManagementBehavior := TOF_Core.GENERIC_MEMORY_MANAGEMENT_BEHAVIOR.STORE_ORIGINAL_REFERENCE_AND_NOT_OWNS_MEMORY
);

__TRY
	comparison := _Actual.CompareTo(otherValue := expectedGeneric);
	isOrdered := (comparison = TOF_Core.COMPARISON_RESULT.FIRST_LESS_THAN_SECOND);
__CATCH
	isOrdered := FALSE;
__ENDTRY

IF NOT isOrdered THEN
	diagnostic := TOF_Core.WideStrings.Concat255(
		"Expected value < ",
		expectedGeneric.AsWString255(),
		", but was: ",
		_Actual.AsWString255()
	);
	fail(defaultMessage := diagnostic);
END_IF

IsLessThan REF= THIS^;
END_METHOD

(*!
<summary>Asserts that the actual value meets the inclusive upper boundary.</summary>
<description>
Uses Core ordering without tolerance. Comparison exceptions record an assertion failure.
The chain message remains available to subsequent assertions.
</description>
<param name="expected">Live variable to compare; ANY does not accept literals or expression results.</param>
*)
METHOD FINAL IsLessThanOrEquals : REFERENCE TO AssertionContext
VAR_INPUT
	expected : ANY;
END_VAR
VAR
	diagnostic : TOF_Core.ERROR_MESSAGE;
	expectedGeneric : TOF_Core.GENERIC_VALUE;
	comparison : TOF_Core.COMPARISON_RESULT;
	isOrdered : BOOL;
END_VAR
expectedGeneric := TOF_Core.GenericValueFactory.FromAny(
	value := expected,
	isObject := FALSE,
	memoryManagementBehavior := TOF_Core.GENERIC_MEMORY_MANAGEMENT_BEHAVIOR.STORE_ORIGINAL_REFERENCE_AND_NOT_OWNS_MEMORY
);

__TRY
	comparison := _Actual.CompareTo(otherValue := expectedGeneric);
	isOrdered := (comparison = TOF_Core.COMPARISON_RESULT.FIRST_LESS_THAN_SECOND)
		OR_ELSE (comparison = TOF_Core.COMPARISON_RESULT.FIRST_EQUAL_TO_SECOND);
__CATCH
	isOrdered := FALSE;
__ENDTRY

IF NOT isOrdered THEN
	diagnostic := TOF_Core.WideStrings.Concat255(
		"Expected value <= ",
		expectedGeneric.AsWString255(),
		", but was: ",
		_Actual.AsWString255()
	);
	fail(defaultMessage := diagnostic);
END_IF

IsLessThanOrEquals REF= THIS^;
END_METHOD

(*!
<summary>Asserts that a typed pointer is non-null. For references assert __ISVALIDREF explicitly.</summary>
<description>
A null pointer or unsupported operand records failure; the chain message remains available.
</description>
*)
METHOD FINAL IsNotNull : REFERENCE TO AssertionContext
IF isNullPointerOrReference() THEN
	fail(defaultMessage := "Expected: non-null object/pointer, but was null (0)");
END_IF

IsNotNull REF= THIS^;
END_METHOD

(*!
<summary>Asserts that a typed pointer is null. For interfaces assert the comparison to zero explicitly.</summary>
<description>
A non-null pointer or unsupported operand records failure; the chain message remains available.
</description>
*)
METHOD FINAL IsNull : REFERENCE TO AssertionContext
IF NOT isNullPointerOrReference() THEN
	fail(defaultMessage := "Expected: null (0), but was non-zero address");
END_IF

IsNull REF= THIS^;
END_METHOD

//! <summary>Reads a typed pointer slot and records unsupported operands as assertion failures.</summary>
METHOD PRIVATE isNullPointerOrReference : BOOL
VAR
	pointerValue : POINTER TO PVOID;
END_VAR
IF _Actual.Address = 0 THEN
	isNullPointerOrReference := TRUE;
	RETURN;
END_IF

IF _Actual.TypeClass = TOF_Core.GENERIC_TYPE_CLASS.POINTER_TO THEN
	pointerValue := _Actual.Address;
	isNullPointerOrReference := (pointerValue^ = 0);
ELSE
	fail(defaultMessage := "Expected a typed pointer. For interfaces or references assert the explicit null predicate.");
END_IF
END_METHOD

(*!
<summary>Asserts that the actual value is a boolean equal to TRUE.</summary>
<description>
A non-Boolean operand or FALSE records failure; the chain message remains available.
</description>
*)
METHOD FINAL IsTrue : REFERENCE TO AssertionContext
VAR
	diagnostic : TOF_Core.ERROR_MESSAGE;
END_VAR
IF _Actual.TypeClass <> TOF_Core.GENERIC_TYPE_CLASS.BOOLEAN OR_ELSE NOT _Actual.AsBool() THEN
	diagnostic := TOF_Core.WideStrings.Concat255(
		"Expected: TRUE, but was: ",
		_Actual.AsWString255()
	);
	fail(defaultMessage := diagnostic);
END_IF

IsTrue REF= THIS^;
END_METHOD

(*!
<summary>Provides the library namespace used in diagnostics.</summary>
<description>
Borrowed read-only reference to the compiler-initialized library namespace; no ownership transfer.
</description>
*)
{attribute 'monitoring' := 'call'}
PROPERTY NamespaceName : REFERENCE TO STRING
GET
NamespaceName REF= CurrentNamespace.Name;
END_GET
END_PROPERTY

(*!
<summary>Asserts exact inequality against a borrowed expected variable.</summary>
<description>
Uses Core value semantics without tolerance. Comparison exceptions record failure, including
for inequality. The message applies to every assertion in the current chain.
</description>
<param name="expected">Live variable to compare; ANY does not accept literals or expression results.</param>
*)
METHOD FINAL NotToBe : REFERENCE TO AssertionContext
VAR_INPUT
	expected : ANY;
END_VAR
VAR
	diagnostic : TOF_Core.ERROR_MESSAGE;
	expectedGeneric : TOF_Core.GENERIC_VALUE;
	areEqual : BOOL;
END_VAR
expectedGeneric := TOF_Core.GenericValueFactory.FromAny(
	value := expected,
	isObject := FALSE,
	memoryManagementBehavior := TOF_Core.GENERIC_MEMORY_MANAGEMENT_BEHAVIOR.STORE_ORIGINAL_REFERENCE_AND_NOT_OWNS_MEMORY
);

__TRY
	areEqual := _Actual.Equals(otherValue := expectedGeneric);
__CATCH
	fail(defaultMessage := "The values could not be compared for equality");
	NotToBe REF= THIS^;
	RETURN;
__ENDTRY

IF areEqual THEN
	diagnostic := TOF_Core.WideStrings.Concat255(
		"Expected value not to be: ",
		expectedGeneric.AsWString255(),
		", but was: ",
		_Actual.AsWString255()
	);
	fail(defaultMessage := diagnostic);
END_IF

NotToBe REF= THIS^;
END_METHOD

(*!
<summary>Prepares one borrowed operand and copies its chain-wide diagnostic prefix.</summary>
<description>
The caller keeps actual storage alive and stable until the immediate chain ends.
Every preparation replaces the message, including an empty message.
</description>
<param name="testCase">Receives failures from this chain.</param>
<param name="actual">Live operand storage borrowed without ownership transfer.</param>
<param name="message">Copied prefix for every assertion in the chain.</param>
*)
METHOD INTERNAL FINAL Prepare : REFERENCE TO AssertionContext
VAR_INPUT
	actual : ANY;
	testCase : ITestCase;
END_VAR
VAR_IN_OUT CONSTANT
	message : WSTRING(255);
END_VAR
_Actual := TOF_Core.GenericValueFactory.FromAny(
	value := actual,
	isObject := FALSE,
	memoryManagementBehavior := TOF_Core.GENERIC_MEMORY_MANAGEMENT_BEHAVIOR.STORE_ORIGINAL_REFERENCE_AND_NOT_OWNS_MEMORY
);
_TestCase := testCase;
_Message := message;

Prepare REF= THIS^;
END_METHOD

(*!
<summary>Reports the byte size of this concrete instance.</summary>
<description>
Uses XSIZEOF on the instance. Does not include separately allocated payloads or prove that an arbitrary
address is valid.
</description>
*)
{attribute 'monitoring' := 'call'}
PROPERTY SelfSize : ULINT
GET
SelfSize := XSIZEOF(THIS^);
END_GET
END_PROPERTY

(*!
<summary>Asserts exact equality against a borrowed expected variable.</summary>
<description>
Uses Core value semantics without tolerance. Comparison exceptions record failure, including
for inequality. The message applies to every assertion in the current chain.
</description>
<param name="expected">Live variable to compare; ANY does not accept literals or expression results.</param>
*)
METHOD FINAL ToBe : REFERENCE TO AssertionContext
VAR_INPUT
	expected : ANY;
END_VAR
VAR
	diagnostic : TOF_Core.ERROR_MESSAGE;
	expectedGeneric : TOF_Core.GENERIC_VALUE;
	areEqual : BOOL;
END_VAR
expectedGeneric := TOF_Core.GenericValueFactory.FromAny(
	value := expected,
	isObject := FALSE,
	memoryManagementBehavior := TOF_Core.GENERIC_MEMORY_MANAGEMENT_BEHAVIOR.STORE_ORIGINAL_REFERENCE_AND_NOT_OWNS_MEMORY
);

__TRY
	areEqual := _Actual.Equals(otherValue := expectedGeneric);
__CATCH
	fail(defaultMessage := "The values could not be compared for equality");
	ToBe REF= THIS^;
	RETURN;
__ENDTRY

IF NOT areEqual THEN
	diagnostic := TOF_Core.WideStrings.Concat255(
		"Expected: ",
		expectedGeneric.AsWString255(),
		", but was: ",
		_Actual.AsWString255()
	);
	fail(defaultMessage := diagnostic);
END_IF

ToBe REF= THIS^;
END_METHOD

(*!
<summary>Asserts that the actual string contains the specified substring.</summary>
<description>
Borrows the actual string and searches by code unit. For STRING_8, searches only if the wide substring
survives conversion to STRING and back to WSTRING. A missing or unrepresentable substring or a non-string
operand records failure without interrupting the callback. The chain message remains available.
</description>
*)
METHOD FINAL ToContain : REFERENCE TO AssertionContext
VAR_INPUT
	substring : WSTRING(255);
END_VAR
VAR
	diagnostic : TOF_Core.ERROR_MESSAGE;
	contains : BOOL;
	convertedSubstring : STRING(255);
END_VAR
IF _Actual.TypeClass = TOF_Core.GENERIC_TYPE_CLASS.STRING_16 THEN
	contains := TOF_Core.WideStrings.Contains(
		stringToSearchIn := _Actual.AsWStringReference(),
		stringToFind := substring
	);
ELSIF _Actual.TypeClass = TOF_Core.GENERIC_TYPE_CLASS.STRING_8 THEN
	convertedSubstring := TO_STRING(substring);

	IF TO_WSTRING(convertedSubstring) = substring THEN
		contains := TOF_Core.Strings.Contains(
			stringToSearchIn := _Actual.AsStringReference(),
			stringToFind := convertedSubstring
		);
	END_IF
END_IF

IF NOT contains THEN
	diagnostic := TOF_Core.WideStrings.Concat255(
		"Expected text to contain '",
		substring,
		"', but was: '",
		_Actual.AsWString255(),
		"'"
	);
	fail(defaultMessage := diagnostic);
END_IF

ToContain REF= THIS^;
END_METHOD

END_FUNCTION_BLOCK

// ---- TestServices.TcPOU
(*
SPDX-FileCopyrightText: © 2026 Oleksandr Tiutyk <trofimich@gmail.com>
SPDX-License-Identifier: MIT
License: https://opensource.org/license/mit
*)

(*!
<summary>Provides internal exception diagnostics and stateless assertion services.</summary>
<description>
Assertion services retain no operands, receiver or diagnostic state between calls. Callers keep borrowed
inputs alive for the call and use each test case only from its owning task without reentry. Failure
reporting propagates receiver exceptions; floating helpers allocate no memory and invoke no callbacks.
</description>
*)

{attribute 'no_explicit_call' := 'do not call this function block directly'}
PROGRAM INTERNAL TestServices
VAR
	{attribute 'hide'} 
	_ClassName : STRING := __POUNAME();
END_VAR

(*!
<summary>Checks canonical floating equality or finite absolute distance without overflowing.</summary>
<description>
Requires canonical binary64 operands and a validated finite nonnegative tolerance. Canonical equality
is accepted first. Zero tolerance does no arithmetic, preserving distinct subnormal representations.
Unequal nonfinite values are never close. Opposite signs use a remaining tolerance budget.
</description>
<param name="actualBits">Canonical actual representation.</param>
<param name="expectedBits">Canonical expected representation.</param>
<param name="tolerance">Validated finite nonnegative absolute distance.</param>
*)
METHOD AreFloatingValuesWithinTolerance : BOOL
VAR_INPUT
	actualBits : ULINT;
	expectedBits : ULINT;
	tolerance : LREAL;
END_VAR
VAR
	actualValue : TOF_Core.LREAL_UNION;
	expectedValue : TOF_Core.LREAL_UNION;
END_VAR
IF actualBits = expectedBits THEN
	AreFloatingValuesWithinTolerance := TRUE;
	RETURN;
END_IF

IF tolerance = TOF_Core.LongReals.ZERO THEN
	RETURN;
END_IF

// The exponent mask isolates binary64 bits 62..52 and rejects remaining nonfinite operands.
IF (actualBits AND TOF_Core.LongReals.EXPONENT_MASK) = TOF_Core.LongReals.EXPONENT_MASK
	OR_ELSE (expectedBits AND TOF_Core.LongReals.EXPONENT_MASK) = TOF_Core.LongReals.EXPONENT_MASK
THEN
	RETURN;
END_IF

actualValue.Raw := actualBits;
expectedValue.Raw := expectedBits;

// Complementing MAGNITUDE_MASK isolates binary64 sign bit 63 to select the safe distance formula.
IF (actualBits AND NOT TOF_Core.LongReals.MAGNITUDE_MASK)
	<> (expectedBits AND NOT TOF_Core.LongReals.MAGNITUDE_MASK)
THEN
	AreFloatingValuesWithinTolerance := ABS(actualValue.Value) <= tolerance
		AND_THEN ABS(expectedValue.Value) <= tolerance - ABS(actualValue.Value);
ELSE
	AreFloatingValuesWithinTolerance := ABS(actualValue.Value - expectedValue.Value) <= tolerance;
END_IF
END_METHOD

//! <summary>Borrows the concrete class name for the lifetime of this instance; callers must not modify it.</summary>
{attribute 'monitoring' := 'call'}
PROPERTY ClassName : REFERENCE TO STRING
GET
ClassName REF= _ClassName;
END_GET
END_PROPERTY

(*!
<summary>Orders canonical floating operands using the Core NaN-first total order.</summary>
<description>
Requires canonical binary64 bits from GetCanonicalRealBits or GetCanonicalLongRealBits. Equal canonical
bits compare equal; NaN precedes every non-NaN value. No comparison evaluates a NaN operand. Other pairs
use native LREAL ordering, including the runtime treatment of subnormal operands.
</description>
<param name="actualBits">Canonical actual representation.</param>
<param name="expectedBits">Canonical expected representation.</param>
*)
METHOD CompareFloatingValues : TOF_Core.COMPARISON_RESULT
VAR_INPUT
	actualBits : ULINT;
	expectedBits : ULINT;
END_VAR
VAR
	actualValue : TOF_Core.LREAL_UNION;
	expectedValue : TOF_Core.LREAL_UNION;
END_VAR
IF actualBits = expectedBits THEN
	CompareFloatingValues := TOF_Core.COMPARISON_RESULT.FIRST_EQUAL_TO_SECOND;
ELSIF actualBits = TOF_Core.LongReals.CANONICAL_NAN_BITS THEN
	CompareFloatingValues := TOF_Core.COMPARISON_RESULT.FIRST_LESS_THAN_SECOND;
ELSIF expectedBits = TOF_Core.LongReals.CANONICAL_NAN_BITS THEN
	CompareFloatingValues := TOF_Core.COMPARISON_RESULT.FIRST_GREATER_THAN_SECOND;
ELSE
	actualValue.Raw := actualBits;
	expectedValue.Raw := expectedBits;

	IF actualValue.Value < expectedValue.Value THEN
		CompareFloatingValues := TOF_Core.COMPARISON_RESULT.FIRST_LESS_THAN_SECOND;
	ELSIF actualValue.Value > expectedValue.Value THEN
		CompareFloatingValues := TOF_Core.COMPARISON_RESULT.FIRST_GREATER_THAN_SECOND;
	ELSE
		CompareFloatingValues := TOF_Core.COMPARISON_RESULT.FIRST_EQUAL_TO_SECOND;
	END_IF
END_IF
END_METHOD

(*!
<summary>Copies a caught exception diagnostic with its callback stage before task cleanup.</summary>
<description>
Borrows the current task's exception only during this call. Returns independent fixed-capacity text;
no exception reference is retained. A failed custom formatter leaves a stage/code fallback.
Terminal allocation failure propagates after the recoverable formatter handler and never becomes a fallback success.
Call only from the owning cyclic task's catch handler; this method neither performs cleanup nor clears the fatal latch.
</description>
<param name="exceptionCode">Native transport code captured by the caller's catch handler.</param>
<param name="stage">Interrupted callback or runner phase included in the copied result.</param>
<param name="catchPointPOUName">POU containing the caller's catch handler.</param>
<param name="catchPointPosition">Source position of the caller's catch handler.</param>
*)
METHOD FormatCaughtException : TOF_Core.ERROR_MESSAGE
VAR_INPUT
	exceptionCode : __SYSTEM.ExceptionCode;
	stage : STRING;
	catchPointPOUName : STRING;
	catchPointPosition : STRING;
END_VAR
VAR
	exception : TOF_Core.IException;
	fallbackMessage : TOF_Core.ERROR_MESSAGE;
	exceptionMessage : TOF_Core.ERROR_MESSAGE;
	diagnostic : TOF_Core.ERROR_MESSAGE;
END_VAR
fallbackMessage := TOF_Core.WideStrings.Concat255(
	TO_WSTRING(stage), ": runtime exception code ", TO_WSTRING(exceptionCode), " (diagnostic unavailable)"
);
FormatCaughtException := fallbackMessage;

// Contain failures from custom exception formatters while preserving the original fallback.
__TRY
	exception := TOF_Core.ExceptionManager.GetLastException(
		exceptionCode := exceptionCode,
		catchPointNamespaceName := CurrentNamespace.Name,
		catchPointPOUName := catchPointPOUName,
		catchPointPosition := catchPointPosition
	);

	IF exception <> 0 THEN
		exceptionMessage := exception.GetMessage(
			showSource := TRUE,
			timestampDisplayMode := TOF_Core.TIMESTAMP_DISPLAY_MODE.HIDDEN
		);
		diagnostic := TO_WSTRING(stage);
		TOF_Core.WideStrings.AppendFit(targetString := diagnostic, sourceString := ": ");
		TOF_Core.WideStrings.AppendFit(targetString := diagnostic, sourceString := exceptionMessage);
		FormatCaughtException := diagnostic;
	END_IF

__CATCH
	FormatCaughtException := fallbackMessage;
__ENDTRY

TOF_Core.DynamicMemoryManager.RaiseIfAllocationFailed();
END_METHOD

(*!
<summary>Maps a LREAL operand to the canonical binary64 assertion representation.</summary>
<description>
Uses LongReals.GetCanonicalBinary64Bits from Core.
Classifies NaN from stored bits and maps all NaNs and signed zeros to Core canonical bits.
Other bit representations are unchanged. No arithmetic, allocation or callback is performed.
</description>
<param name="value">Typed operand copied for this call.</param>
*)
METHOD GetCanonicalLongRealBits : ULINT
VAR_INPUT
	value : LREAL;
END_VAR
GetCanonicalLongRealBits := TOF_Core.LongReals.GetCanonicalBinary64Bits(value := value);
END_METHOD

(*!
<summary>Maps a REAL operand to the canonical binary64 assertion representation.</summary>
<description>
Uses Reals.GetCanonicalBinary64Bits from Core.
Classifies NaN before arithmetic or widening, maps all NaNs and signed zeros to Core canonical bits.
Other REAL values widen to LREAL using the runtime floating configuration. Owns no resources.
</description>
<param name="value">Typed operand copied for this call.</param>
*)
METHOD GetCanonicalRealBits : ULINT
VAR_INPUT
	value : REAL;
END_VAR
GetCanonicalRealBits := TOF_Core.Reals.GetCanonicalBinary64Bits(value := value);
END_METHOD

(*!
<summary>Checks whether an absolute tolerance is finite and nonnegative.</summary>
<description>
Rejects NaN and infinity from the stored exponent before arithmetic. Returns FALSE without reporting
failure; the calling typed context reports the invalid argument with its current chain message.
</description>
<param name="tolerance">Absolute comparison distance; zero requests canonical equality.</param>
*)
METHOD IsValidFloatingTolerance : BOOL
VAR_INPUT
	tolerance : LREAL;
END_VAR
VAR
	bits : TOF_Core.LREAL_UNION;
END_VAR
bits.Value := tolerance;

// Binary64 exponent bits 62..52 are all set for infinity and NaN.
IsValidFloatingTolerance := (bits.Raw AND TOF_Core.LongReals.EXPONENT_MASK) <> TOF_Core.LongReals.EXPONENT_MASK
	AND_THEN tolerance >= TOF_Core.LongReals.ZERO;
END_METHOD

//! <summary>Borrows the compiler-initialized namespace; callers must not modify the returned reference.</summary>
{attribute 'monitoring' := 'call'}
PROPERTY NamespaceName : REFERENCE TO STRING
GET
NamespaceName REF= CurrentNamespace.Name;
END_GET
END_PROPERTY

(*!
<summary>Reports a failed predicate with the copied chain prefix.</summary>
<description>
A missing receiver raises DataMemberNotSpecifiedException. A whitespace-only prefix is omitted.
The receiver decides whether to retain the diagnostic; callback exceptions propagate. No input is retained.
</description>
<param name="testCase">Borrowed failure receiver.</param>
<param name="message">Chain prefix copied by the calling context.</param>
<param name="sourceClassName">Calling context class used for a missing-receiver diagnostic.</param>
<param name="defaultMessage">Assertion diagnostic borrowed for this call.</param>
*)
METHOD ReportAssertionFailure
VAR_INPUT
	testCase : ITestCase;
	message : WSTRING(255);
	sourceClassName : STRING;
END_VAR
VAR_IN_OUT CONSTANT
	defaultMessage : TOF_Core.ERROR_MESSAGE;
END_VAR
VAR
	diagnostic : TOF_Core.ERROR_MESSAGE;
END_VAR
IF testCase = 0 THEN
	TOF_Core.Exceptions.ThrowDataMemberNotSpecified(
		sourceNamespaceName := NamespaceName,
		sourceClassName := sourceClassName,
		sourcePOUName := __POUNAME(),
		sourcePosition := __POSITION(),
		dataMemberName := '_TestCase'
	);
END_IF

IF TOF_Core.WideStrings.IsNullOrWhiteSpace(stringToCheck := message) THEN
	testCase.RecordFailure(message := defaultMessage);
ELSE
	diagnostic := message;
	TOF_Core.WideStrings.AppendFit(targetString := diagnostic, sourceString := ": ");
	TOF_Core.WideStrings.AppendFit(targetString := diagnostic, sourceString := defaultMessage);
	testCase.RecordFailure(message := diagnostic);
END_IF
END_METHOD

END_PROGRAM

// ---- Internal/CurrentNamespace.TcPOU
(*
SPDX-FileCopyrightText: © 2026 Oleksandr Tiutyk <trofimich@gmail.com>
SPDX-License-Identifier: MIT
License: https://opensource.org/license/mit
*)

(*!
<summary>Exposes the compiler-initialized namespace of the Testing library.</summary>
<description>Static internal storage; Name is a borrowed read-only view and requires no cyclic execution.</description>
*)

{attribute 'no_explicit_call' := 'do not call this POU directly'}
PROGRAM INTERNAL CurrentNamespace
VAR
	{attribute 'hide'} 
	_NamespaceExtractor : NamespaceExtractor;
	_ClassName : STRING := __POUNAME();
END_VAR

(*!
<summary>Returns the compiler-initialized library namespace.</summary>
<description>Borrowed read-only reference to static storage. Do not modify it through the reference.</description>
*)
{attribute 'monitoring' := 'call'}
PROPERTY Name : REFERENCE TO STRING
GET
Name REF= _NamespaceExtractor.CurrentNamespace;
END_GET
END_PROPERTY

(*!
<summary>Borrows the concrete metadata provider name for its lifetime.</summary>
<description>Borrowed read-only storage; callers must not modify it.</description>
*)
{attribute 'monitoring' := 'call'}
PROPERTY ClassName : REFERENCE TO STRING
GET
ClassName REF= _ClassName;
END_GET
END_PROPERTY

(*!
<summary>Borrows the compiler-initialized library namespace.</summary>
<description>Borrowed read-only storage; callers must not modify it.</description>
*)
{attribute 'monitoring' := 'call'}
PROPERTY NamespaceName : REFERENCE TO STRING
GET
NamespaceName REF= _NamespaceExtractor.CurrentNamespace;
END_GET
END_PROPERTY

END_PROGRAM

// ---- Internal/NamespaceExtractor.TcPOU
(*
SPDX-FileCopyrightText: © 2026 Oleksandr Tiutyk <trofimich@gmail.com>
SPDX-License-Identifier: MIT
License: https://opensource.org/license/mit
*)

(*!
<summary>Obtains the library namespace through the init_namespace attribute.</summary>
<description>
Internal static metadata holder. Its output is initialized by TwinCAT rather than by cyclic execution.
</description>
*)

{attribute 'no_explicit_call' := 'do not call this function block directly'}
FUNCTION_BLOCK INTERNAL NamespaceExtractor
VAR_OUTPUT
	{attribute 'init_namespace'} 
	CurrentNamespace : STRING;	
END_VAR

END_FUNCTION_BLOCK

// ---- TestElements/Tests/TestCase.TcPOU
(*
SPDX-FileCopyrightText: © 2026 Oleksandr Tiutyk <trofimich@gmail.com>
SPDX-License-Identifier: MIT
License: https://opensource.org/license/mit
*)

(*!
<summary>Owns the lifecycle and copied diagnostic of one leaf test.</summary>
<description>
BeforeTest runs once; ExecuteTest runs according to the concrete single-cycle or multi-cycle strategy.
AfterTest runs once after normal completion, assertion failure, deadline or a caught scenario exception,
including failed preparation. Teardown must tolerate partially prepared resources. Assertions record failure
without interrupting the remaining statements of the callback. The first failure diagnostic is retained, including copied exception text/source and callback stage.
A failing exception formatter produces a stage/code fallback without replacing an earlier failure.
Exceptions from scenario hooks become one failed leaf result; catches do not roll back user side effects.
Terminal OOM propagates outside recoverable handlers and stops normal execution; teardown is not promised then.
Throwing callbacks must not use method-local resource-owning FBs that require stack unwinding.
Path-provider and reporter exceptions propagate after terminal state is committed and the stored reporter reference
is cleared. Completed callbacks are never retried.
</description>
*)

{attribute 'no_explicit_call' := 'do not call this function block directly'}
FUNCTION_BLOCK ABSTRACT TestCase EXTENDS TestElement IMPLEMENTS ITestCase
VAR
	//! <summary>Assertions bound to this case; finish one chain before starting another.</summary>
	_Assert : Assertions;	
	_Outcome : TEST_OUTCOME;
	_FailureMessage : TOF_Core.ERROR_MESSAGE;
	_Elapsed : LTIME;
	_CycleCount : UDINT;
END_VAR

(*!
<summary>Cleans up this scenario once, including after preparation or body failure.</summary>
*)
METHOD PROTECTED AfterTest
END_METHOD

(*!
<summary>Borrows the assertions bound to this running test case.</summary>
<description>Complete one immediate chain at a time; do not retain it or mutate the provider.</description>
*)
{attribute 'monitoring' := 'call'}
PROPERTY FINAL Assert : REFERENCE TO Assertions
GET
Assert REF= _Assert;
END_GET
END_PROPERTY

(*!
<summary>Prepares this scenario once per run; teardown must handle partial preparation.</summary>
*)
METHOD PROTECTED BeforeTest
END_METHOD

(*!
<summary>Counts scheduling cycles, including a deadline cycle; saturates at the UDINT maximum.</summary>
*)
{attribute 'monitoring' := 'call'}
PROPERTY FINAL CycleCount : UDINT
GET
CycleCount := _CycleCount;
END_GET
END_PROPERTY

(*!
<summary>Reports nominal time since the first scheduling cycle, initially zero.</summary>
*)
{attribute 'monitoring' := 'call'}
PROPERTY FINAL Elapsed : TIME
GET
Elapsed := TO_TIME(_Elapsed);
END_GET
END_PROPERTY

(*!
<summary>Schedules one leaf cycle and commits one result after teardown.</summary>
<description>
Scenario exceptions are converted to FAILED so the containing sequence can continue. Completion clears the
stored reporter reference before path lookup and result delivery. Exceptions from either callback propagate.
</description>
*)
// Manual stack estimate for TwinCAT. Reassess if callbacks or test workloads change.
{attribute 'estimated-stack-usage' := '16384'}
METHOD FINAL Execute
VAR
	resultReporter : ITestReporter;
	groupPath : WSTRING(255);
	exceptionCode : __SYSTEM.ExceptionCode;
	cycleResult : TEST_CYCLE_RESULT;
END_VAR
IF IsFinished THEN
	RETURN;
END_IF

IF _State = TEST_ELEMENT_STATE.READY THEN
	_State := TEST_ELEMENT_STATE.RUNNING;
	_Outcome := TEST_OUTCOME.RUNNING;
	_CycleCount := 1;
	
	_Assert.Bind(testCase := THIS^);

	__TRY
		BeforeTest();
	__CATCH(exceptionCode)
		recordRuntimeException(
			exceptionCode := exceptionCode,
			stage := 'BeforeTest',
			catchPointPOUName := __POUNAME(),
			catchPointPosition := __POSITION()
		);
	__ENDTRY

	TOF_Core.DynamicMemoryManager.RaiseIfAllocationFailed();
ELSE
	IF _CycleCount < TOF_Core.UnsignedInt32.MAX_VALUE THEN
		_CycleCount := _CycleCount + 1;
	END_IF

	_Elapsed := _Elapsed + TOF_Core.System.GetTaskCycleTime();
END_IF

_Duration := _Duration + TOF_Core.System.GetTaskCycleTime();

IF _Outcome <> TEST_OUTCOME.FAILED THEN
	__TRY
		cycleResult := RunCycle();
	__CATCH(exceptionCode)
		recordRuntimeException(
			exceptionCode := exceptionCode,
			stage := 'ExecuteTest',
			catchPointPOUName := __POUNAME(),
			catchPointPosition := __POSITION()
		);
	__ENDTRY
END_IF

TOF_Core.DynamicMemoryManager.RaiseIfAllocationFailed();

IF cycleResult <> TEST_CYCLE_RESULT.DONE AND_THEN _Outcome <> TEST_OUTCOME.FAILED THEN
	RETURN;
END_IF

__TRY
	AfterTest();
__CATCH(exceptionCode)
	recordRuntimeException(
		exceptionCode := exceptionCode,
		stage := 'AfterTest',
		catchPointPOUName := __POUNAME(),
		catchPointPosition := __POSITION()
	);
__ENDTRY

TOF_Core.DynamicMemoryManager.RaiseIfAllocationFailed();

IF _Outcome = TEST_OUTCOME.FAILED THEN
	_FailedCount := 1;
ELSE
	_Outcome := TEST_OUTCOME.PASSED;
	_PassedCount := 1;
END_IF

resultReporter := _Reporter;
_Reporter := 0;
_State := TEST_ELEMENT_STATE.COMPLETED;

IF resultReporter <> 0 THEN
	IF _Parent <> 0 THEN
		groupPath := _Parent.GetPath();
	END_IF

	resultReporter.ReportTestCaseResult(
		groupPath := groupPath,
		testName := _Name,
		outcome := _Outcome,
		duration := Duration,
		message := _FailureMessage
	);
END_IF
END_METHOD

(*!
<summary>Borrows the first copied failure diagnostic.</summary>
*)
{attribute 'monitoring' := 'call'}
PROPERTY FINAL FailureMessage : REFERENCE TO TOF_Core.ERROR_MESSAGE
GET
FailureMessage REF= _FailureMessage;
END_GET
END_PROPERTY

(*!
<summary>Reports this leaf execution outcome.</summary>
*)
{attribute 'monitoring' := 'call'}
PROPERTY FINAL Outcome : TEST_OUTCOME
GET
Outcome := _Outcome;
END_GET
END_PROPERTY

(*!
<summary>Copies the first failure while the case is running.</summary>
<description>
Does not throw for a test failure, interrupt the current callback, or change an already completed result.
</description>
*)
METHOD FINAL RecordFailure
VAR_IN_OUT CONSTANT
	message : TOF_Core.ERROR_MESSAGE;
END_VAR
IF _State <> TEST_ELEMENT_STATE.RUNNING OR_ELSE _Outcome = TEST_OUTCOME.FAILED THEN
	RETURN;
END_IF

_Outcome := TEST_OUTCOME.FAILED;
_FailureMessage := message;
END_METHOD

(*!
<summary>Copies a caught hook exception as a leaf failure without retaining its object.</summary>
<description>Preserves an earlier failure and forwards the actual catch location to diagnostic formatting.</description>
*)
METHOD PRIVATE recordRuntimeException
VAR_INPUT
	exceptionCode : __SYSTEM.ExceptionCode;
	stage : STRING;
	catchPointPOUName : STRING;
	catchPointPosition : STRING;
END_VAR
VAR
	diagnostic : TOF_Core.ERROR_MESSAGE;
END_VAR
IF _Outcome = TEST_OUTCOME.FAILED THEN
	RETURN;
END_IF

diagnostic := TestServices.FormatCaughtException(
	exceptionCode := exceptionCode,
	stage := stage,
	catchPointPOUName := catchPointPOUName,
	catchPointPosition := catchPointPosition
);
RecordFailure(message := diagnostic);
END_METHOD

(*!
<summary>Prepares fresh leaf observations without running scenario hooks.</summary>
<description>
Does not run teardown or release user resources. Call only at the lifecycle boundaries in ITestElement.
The reporter is borrowed until completion; no locks or cross-task transfer are provided.
Clears this case's outcome, diagnostic and nominal timing after common state is reset.
</description>
*)
METHOD FINAL Reset
VAR_INPUT
	reporter : ITestReporter;
END_VAR
SUPER^.Reset(reporter := reporter);

_Outcome := TEST_OUTCOME.NOT_RUN;
_FailureMessage := "";
_Elapsed := LTIME#0NS;
_CycleCount := 0;
END_METHOD

(*!
<summary>Applies the concrete scheduling strategy and returns whether the cycle finished the body.</summary>
*)
METHOD PROTECTED ABSTRACT RunCycle : TEST_CYCLE_RESULT
END_METHOD

(*!
<summary>Counts this single scenario regardless of execution state or outcome.</summary>
*)
{attribute 'monitoring' := 'call'}
PROPERTY FINAL TestCount : TOF_Core.DINT_LENGTH
GET
TestCount := 1;
END_GET
END_PROPERTY

END_FUNCTION_BLOCK

// ---- TestElements/TestElement.TcPOU
(*
SPDX-FileCopyrightText: © 2026 Oleksandr Tiutyk <trofimich@gmail.com>
SPDX-License-Identifier: MIT
License: https://opensource.org/license/mit
*)

(*!
<summary>Shares names, computed paths, lifecycle observations and borrowed tree links between test elements.</summary>
<description>
Construction copies the display name and assigned parent without invoking callbacks or inspecting the tree.
No automatic registration or deletion of children or reporters occurs. Parent links are fixed structural assignments,
not allocation ownership. Do not copy instances by value or change configuration during execution.
Descendants implement execution, reset their own state and supply the configured leaf count.
Reset is not cancellation; recover resources explicitly before resetting an externally aborted tree.
Concrete descendants implement the Object metadata properties for their own class, namespace and instance size.
Inherited Object equality and hashing use instance identity unless a descendant overrides both consistently.
</description>
*)

{attribute 'no_explicit_call' := 'do not call this function block directly'}
FUNCTION_BLOCK ABSTRACT TestElement EXTENDS TOF_Core.Object IMPLEMENTS ITestElement
VAR
	{attribute 'hide'} 
	_Name : WSTRING;
	
	{attribute 'hide'} 
	_Parent : ITestElement;

	{attribute 'hide'} 
	_Reporter : ITestReporter;

	{attribute 'hide'} 
	_State : TEST_ELEMENT_STATE;

	{attribute 'hide'} 
	_PassedCount : TOF_Core.DINT_LENGTH;
	{attribute 'hide'} 
	_FailedCount : TOF_Core.DINT_LENGTH;
	{attribute 'hide'} 
	_SkippedCount : TOF_Core.DINT_LENGTH;
	
	{attribute 'hide'} 
	_Duration : LTIME;
END_VAR

(*!
<summary>Reports nominal scheduled duration, not CPU execution time.</summary>
*)
{attribute 'monitoring' := 'call'}
PROPERTY FINAL Duration : TIME
GET
Duration := TO_TIME(_Duration);
END_GET
END_PROPERTY

(*!
<summary>Advances the concrete element once; descendants preserve the ITestElement lifecycle.</summary>
*)
METHOD ABSTRACT Execute
END_METHOD

(*!
<summary>Counts failed leaves.</summary>
*)
{attribute 'monitoring' := 'call'}
PROPERTY FINAL FailedCount : TOF_Core.DINT_LENGTH
GET
FailedCount := _FailedCount;
END_GET
END_PROPERTY

(*!
<summary>Copies the display name and fixed parent without invoking overridable code.</summary>
<description>
Copies the borrowed parent without calling it or validating topology. Roots explicitly pass zero.
The parent must remain alive throughout this element's lifetime; construction never raises exceptions.
</description>
<param name="name">Copied display name of at most 80 wide characters; longer input is truncated by IEC conversion.</param>
<param name="parent">Assigned group for the instance lifetime, or zero for a root.</param>
*)
METHOD FB_init : BOOL
VAR_INPUT
	bInitRetains : BOOL; // TRUE: the retain variables are initialized (reset warm / reset cold)
	bInCopyCode : BOOL; // TRUE: the instance will be copied to the copy code afterward (online change)
	name : WSTRING;
	parent : ITestElement;
END_VAR
_Name := name;
_Parent := parent;
END_METHOD

(*!
<summary>Builds the full display path from the root through this element.</summary>
<description>
Joins nonempty names with '/', including this element's name. A nameless root returns an empty path.
The result is a copied WSTRING bounded to 255 characters; overflow preserves the root prefix and ends with an ellipsis.
Reads the live Parent and Name properties without caching or changing the tree. All providers must remain alive
and stable during the call; use only in the owning task without reentry. Can be called before Reset.
A cyclic Parent chain raises StandardException to prevent an endless traversal. Provider exceptions propagate;
no element state or ownership is changed. Valid traversal uses fixed local strings without recursion or heap allocation.
</description>
*)
METHOD FINAL GetPath : WSTRING(255)
VAR
	ancestor : ITestElement;
	slowAncestor : ITestElement;
	fastAncestor : ITestElement;
	descendantPath : WSTRING(255);
END_VAR
ancestor := THIS^;
slowAncestor := ancestor;
fastAncestor := ancestor;

// Reject a cyclic parent chain before constructing any path or invoking another GetPath.
WHILE fastAncestor <> 0 DO
	fastAncestor := fastAncestor.Parent;

	IF fastAncestor = 0 THEN
		EXIT;
	END_IF

	fastAncestor := fastAncestor.Parent;
	slowAncestor := slowAncestor.Parent;

	IF fastAncestor <> 0 AND_THEN fastAncestor = slowAncestor THEN
		TOF_Core.Exceptions.ThrowStandard(
			sourceNamespaceName := NamespaceName,
			sourceClassName := ClassName,
			sourcePOUName := __POUNAME(),
			sourcePosition := __POSITION(),
			message := "The assigned parent chain contains a cycle"
		);
	END_IF
END_WHILE

// Prepending each nonempty ancestor preserves the root prefix when the bounded path overflows.
WHILE ancestor <> 0 DO
	IF ancestor.Name <> "" THEN
		descendantPath := GetPath;
		GetPath := "";
		TOF_Core.WideStrings.AppendFit(targetString := GetPath, sourceString := ancestor.Name);

		IF descendantPath <> "" THEN
			TOF_Core.WideStrings.AppendFit(targetString := GetPath, sourceString := "/");
			TOF_Core.WideStrings.AppendFit(targetString := GetPath, sourceString := descendantPath);
		END_IF
	END_IF

	ancestor := ancestor.Parent;
END_WHILE
END_METHOD

(*!
<summary>Reports terminal completion.</summary>
*)
{attribute 'monitoring' := 'call'}
PROPERTY FINAL IsFinished : BOOL
GET
IsFinished := _State = TEST_ELEMENT_STATE.COMPLETED;
END_GET
END_PROPERTY

(*!
<summary>Reports an active run.</summary>
*)
{attribute 'monitoring' := 'call'}
PROPERTY FINAL IsRunning : BOOL
GET
IsRunning := _State = TEST_ELEMENT_STATE.RUNNING;
END_GET
END_PROPERTY

(*!
<summary>Borrows the display name through the INamed property signature.</summary>
<description>
The reference aliases the constructor-copied name of at most 80 wide characters and remains valid while this element lives.
Callers must not modify the returned reference; no ownership is transferred.
</description>
*)
{attribute 'monitoring' := 'call'}
PROPERTY FINAL Name : REFERENCE TO WSTRING
GET
Name REF= _Name;
END_GET
END_PROPERTY

(*!
<summary>Returns the parent assigned at construction; roots have no parent.</summary>
<description>Borrowed lifetime association, not a registration or allocation-ownership transfer.
The value remains unchanged across Reset and execution; the parent must outlive this element.</description>
*)
{attribute 'monitoring' := 'call'}
PROPERTY FINAL Parent : ITestElement
GET
Parent := _Parent;
END_GET
END_PROPERTY

(*!
<summary>Counts passed leaves.</summary>
*)
{attribute 'monitoring' := 'call'}
PROPERTY FINAL PassedCount : TOF_Core.DINT_LENGTH
GET
PassedCount := _PassedCount;
END_GET
END_PROPERTY

(*!
<summary>Reports nominal scheduled duration, not CPU execution time.</summary>
*)
{attribute 'monitoring' := 'call'}
PROPERTY FINAL Reporter : ITestReporter
GET
Reporter := _Reporter;
END_GET
END_PROPERTY

(*!
<summary>Clears common execution observations and borrows the reporter for a fresh run.</summary>
<description>
Does not run teardown or release user resources. Call only at the lifecycle boundaries in ITestElement.
The reporter is borrowed until completion; no locks or cross-task transfer are provided.
Derived reset failures propagate and can leave a partially reset tree; the runner aborts startup.
Custom element overrides reset their own observations and call SUPER^.Reset with the same reporter.
The base implementation resets only common observations; there is no OnReset callback.
</description>
*)
METHOD Reset
VAR_INPUT
	reporter : ITestReporter;
END_VAR
_Reporter := reporter;
_State := TEST_ELEMENT_STATE.READY;
_PassedCount := 0;
_FailedCount := 0;
_SkippedCount := 0;
_Duration := LTIME#0NS;
END_METHOD

(*!
<summary>Counts skipped leaves.</summary>
*)
{attribute 'monitoring' := 'call'}
PROPERTY FINAL SkippedCount : TOF_Core.DINT_LENGTH
GET
SkippedCount := _SkippedCount;
END_GET
END_PROPERTY

(*!
<summary>Reports nominal scheduled duration, not CPU execution time.</summary>
*)
{attribute 'monitoring' := 'call'}
PROPERTY FINAL State : TEST_ELEMENT_STATE
GET
State := _State;
END_GET
END_PROPERTY

(*!
<summary>Provides the leaf count defined by ITestElement.TestCount.</summary>
*)
{attribute 'monitoring' := 'call'}
PROPERTY ABSTRACT TestCount : TOF_Core.DINT_LENGTH
GET
END_GET
END_PROPERTY

END_FUNCTION_BLOCK

// ---- Assertions/TypedContexts/BoolAssertionContext.TcPOU
(*
SPDX-FileCopyrightText: © 2026 Oleksandr Tiutyk <trofimich@gmail.com>
SPDX-License-Identifier: MIT
License: https://opensource.org/license/mit
*)

(*!
<summary>Provides fluent assertions on a copied BOOL value.</summary>
<description>
Copies actual into persistent instance storage before the entry method returns; literals and expression
results therefore remain valid throughout the immediate chain. Owns no heap allocation or pointed-to resource.
The message prefixes every failure until the next preparation. Finish one chain before starting another on
the owning Assertions provider. Use only from the owning test callback on one task, without reentry.
Obtain this context from the owning provider; direct unprepared use is unsupported.
Expected arguments use the declared IEC type; ordinary compiler conversions happen before comparison.
This context does not depend on another assertion context.
Object metadata is available before preparation; inherited equality compares instance identity.
</description>
*)

{attribute 'no_explicit_call' := 'do not call this function block directly'}
FUNCTION_BLOCK BoolAssertionContext EXTENDS TOF_Core.Object
VAR_STAT
	{attribute 'hide'}
	_ClassName : STRING := __POUNAME();
END_VAR
VAR
	_Actual : BOOL;
	_TestCase : ITestCase;
	_Message : WSTRING(255);
END_VAR

(*!
<summary>Provides the implementation class name.</summary>
<description>
Borrowed read-only reference to compiler-initialized storage, valid throughout the instance lifetime.
Do not modify the returned reference; no ownership is transferred.
</description>
*)
{attribute 'monitoring' := 'call'}
PROPERTY ClassName : REFERENCE TO STRING
GET
ClassName REF= _ClassName;
END_GET
END_PROPERTY

(*!
<summary>Asserts that the actual Boolean value is FALSE.</summary>
<description>
Records failure without interrupting the callback; preserves the chain message.
</description>
*)
METHOD FINAL IsFalse : REFERENCE TO BoolAssertionContext
IF _Actual THEN
	failComparison(expected := FALSE, expectation := "Expected: ");
END_IF

IsFalse REF= THIS^;
END_METHOD

(*!
<summary>Asserts that the actual Boolean value is TRUE.</summary>
<description>
Records failure without interrupting the callback; preserves the chain message.
</description>
*)
METHOD FINAL IsTrue : REFERENCE TO BoolAssertionContext
IF NOT _Actual THEN
	failComparison(expected := TRUE, expectation := "Expected: ");
END_IF

IsTrue REF= THIS^;
END_METHOD

(*!
<summary>Provides the library namespace.</summary>
<description>
Borrowed read-only reference to the compiler-initialized namespace, valid throughout the instance lifetime.
Do not modify the returned reference; no ownership is transferred.
</description>
*)
{attribute 'monitoring' := 'call'}
PROPERTY NamespaceName : REFERENCE TO STRING
GET
NamespaceName REF= CurrentNamespace.Name;
END_GET
END_PROPERTY

(*!
<summary>Asserts inequality with the expected value.</summary>
<description>
Records failure without interrupting the callback; preserves the message for the rest of the chain.
</description>
<param name="expected">Expected value converted by the compiler to BOOL.</param>
*)
METHOD FINAL NotToBe : REFERENCE TO BoolAssertionContext
VAR_INPUT
	expected : BOOL;
END_VAR
IF _Actual = expected THEN
	failComparison(
		expected := expected,
		expectation := "Expected value not to be: "
	);
END_IF

NotToBe REF= THIS^;
END_METHOD

(*!
<summary>Copies the actual operand and replaces the chain-wide message.</summary>
<description>
Called by the owning Assertions provider after it verifies the running test case.
No pointer to this method's input storage is retained. The receiver is borrowed until the next preparation;
the owning provider keeps it alive throughout the immediate chain.
</description>
<param name="actual">Value copied into this context.</param>
<param name="testCase">Borrowed failure receiver for the immediate chain.</param>
<param name="message">Copied diagnostic prefix, including empty to clear the previous prefix.</param>
*)
METHOD INTERNAL FINAL Prepare
VAR_INPUT
	actual : BOOL;
	testCase : ITestCase;
END_VAR
VAR_IN_OUT CONSTANT
	message : WSTRING(255);
END_VAR
_Actual := actual;
_TestCase := testCase;
_Message := message;
END_METHOD

(*!
<summary>Reports the byte size of this concrete instance.</summary>
<description>
Includes inline fields and nested instances, but excludes separately allocated payloads.
Obtaining the size does not transfer ownership or validate an arbitrary address.
</description>
*)
{attribute 'monitoring' := 'call'}
PROPERTY SelfSize : ULINT
GET
SelfSize := XSIZEOF(THIS^);
END_GET
END_PROPERTY

(*!
<summary>Asserts equality with the expected value.</summary>
<description>
Records failure without interrupting the callback; preserves the message for the rest of the chain.
</description>
<param name="expected">Expected value converted by the compiler to BOOL.</param>
*)
METHOD FINAL ToBe : REFERENCE TO BoolAssertionContext
VAR_INPUT
	expected : BOOL;
END_VAR
IF _Actual <> expected THEN
	failComparison(
		expected := expected,
		expectation := "Expected: "
	);
END_IF

ToBe REF= THIS^;
END_METHOD

(*!
<summary>Formats a failed typed predicate and reports it with the chain message.</summary>
<description>
Does not change operands or chain state. The receiver retains its first failure. Reporting exceptions
propagate to the enclosing test callback handler; an unprepared receiver is a configuration error.
</description>
<param name="expected">Typed expected operand used only for this diagnostic.</param>
<param name="expectation">Prefix identifying the failed predicate.</param>
*)
METHOD PRIVATE failComparison
VAR_INPUT
	expected : BOOL;
	expectation : WSTRING(40);
END_VAR
VAR
	actualText : WSTRING(255);
	expectedText : WSTRING(255);
	diagnostic : TOF_Core.ERROR_MESSAGE;
END_VAR
actualText := TO_WSTRING(_Actual);
expectedText := TO_WSTRING(expected);

diagnostic := TOF_Core.WideStrings.Concat255(
	expectation,
	expectedText,
	", but was: ",
	actualText
);

TestServices.ReportAssertionFailure(
	testCase := _TestCase,
	message := _Message,
	sourceClassName := ClassName,
	defaultMessage := diagnostic
);
END_METHOD

END_FUNCTION_BLOCK

// ---- Assertions/TypedContexts/SIntAssertionContext.TcPOU
(*
SPDX-FileCopyrightText: © 2026 Oleksandr Tiutyk <trofimich@gmail.com>
SPDX-License-Identifier: MIT
License: https://opensource.org/license/mit
*)

(*!
<summary>Provides fluent assertions on a copied SINT value.</summary>
<description>
Copies actual into persistent instance storage before the entry method returns; literals and expression
results therefore remain valid throughout the immediate chain. Owns no heap allocation or pointed-to resource.
The message prefixes every failure until the next preparation. Finish one chain before starting another on
the owning Assertions provider. Use only from the owning test callback on one task, without reentry.
Obtain this context from the owning provider; direct unprepared use is unsupported.
Expected arguments use the declared IEC type; ordinary compiler conversions happen before comparison.
This context does not depend on another assertion context.
Object metadata is available before preparation; inherited equality compares instance identity.
</description>
*)

{attribute 'no_explicit_call' := 'do not call this function block directly'}
FUNCTION_BLOCK SIntAssertionContext EXTENDS TOF_Core.Object
VAR_STAT
	{attribute 'hide'}
	_ClassName : STRING := __POUNAME();
END_VAR
VAR
	_Actual : SINT;
	_TestCase : ITestCase;
	_Message : WSTRING(255);
END_VAR

(*!
<summary>Provides the implementation class name.</summary>
<description>
Borrowed read-only reference to compiler-initialized storage, valid throughout the instance lifetime.
Do not modify the returned reference; no ownership is transferred.
</description>
*)
{attribute 'monitoring' := 'call'}
PROPERTY ClassName : REFERENCE TO STRING
GET
ClassName REF= _ClassName;
END_GET
END_PROPERTY

(*!
<summary>Asserts that the actual value is strictly greater than expected.</summary>
<description>
Records failure without interrupting the callback; preserves the message for the rest of the chain.
</description>
<param name="expected">Expected value converted by the compiler to SINT.</param>
*)
METHOD FINAL IsGreaterThan : REFERENCE TO SIntAssertionContext
VAR_INPUT
	expected : SINT;
END_VAR
IF _Actual <= expected THEN
	failComparison(
		expected := expected,
		expectation := "Expected value > "
	);
END_IF

IsGreaterThan REF= THIS^;
END_METHOD

(*!
<summary>Asserts that the actual value meets the inclusive lower boundary.</summary>
<description>
Records failure without interrupting the callback; preserves the message for the rest of the chain.
</description>
<param name="expected">Expected value converted by the compiler to SINT.</param>
*)
METHOD FINAL IsGreaterThanOrEquals : REFERENCE TO SIntAssertionContext
VAR_INPUT
	expected : SINT;
END_VAR
IF _Actual < expected THEN
	failComparison(
		expected := expected,
		expectation := "Expected value >= "
	);
END_IF

IsGreaterThanOrEquals REF= THIS^;
END_METHOD

(*!
<summary>Asserts that the actual value is strictly less than expected.</summary>
<description>
Records failure without interrupting the callback; preserves the message for the rest of the chain.
</description>
<param name="expected">Expected value converted by the compiler to SINT.</param>
*)
METHOD FINAL IsLessThan : REFERENCE TO SIntAssertionContext
VAR_INPUT
	expected : SINT;
END_VAR
IF _Actual >= expected THEN
	failComparison(
		expected := expected,
		expectation := "Expected value < "
	);
END_IF

IsLessThan REF= THIS^;
END_METHOD

(*!
<summary>Asserts that the actual value meets the inclusive upper boundary.</summary>
<description>
Records failure without interrupting the callback; preserves the message for the rest of the chain.
</description>
<param name="expected">Expected value converted by the compiler to SINT.</param>
*)
METHOD FINAL IsLessThanOrEquals : REFERENCE TO SIntAssertionContext
VAR_INPUT
	expected : SINT;
END_VAR
IF _Actual > expected THEN
	failComparison(
		expected := expected,
		expectation := "Expected value <= "
	);
END_IF

IsLessThanOrEquals REF= THIS^;
END_METHOD

(*!
<summary>Provides the library namespace.</summary>
<description>
Borrowed read-only reference to the compiler-initialized namespace, valid throughout the instance lifetime.
Do not modify the returned reference; no ownership is transferred.
</description>
*)
{attribute 'monitoring' := 'call'}
PROPERTY NamespaceName : REFERENCE TO STRING
GET
NamespaceName REF= CurrentNamespace.Name;
END_GET
END_PROPERTY

(*!
<summary>Asserts inequality with the expected value.</summary>
<description>
Records failure without interrupting the callback; preserves the message for the rest of the chain.
</description>
<param name="expected">Expected value converted by the compiler to SINT.</param>
*)
METHOD FINAL NotToBe : REFERENCE TO SIntAssertionContext
VAR_INPUT
	expected : SINT;
END_VAR
IF _Actual = expected THEN
	failComparison(
		expected := expected,
		expectation := "Expected value not to be: "
	);
END_IF

NotToBe REF= THIS^;
END_METHOD

(*!
<summary>Copies the actual operand and replaces the chain-wide message.</summary>
<description>
Called by the owning Assertions provider after it verifies the running test case.
No pointer to this method's input storage is retained. The receiver is borrowed until the next preparation;
the owning provider keeps it alive throughout the immediate chain.
</description>
<param name="actual">Value copied into this context.</param>
<param name="testCase">Borrowed failure receiver for the immediate chain.</param>
<param name="message">Copied diagnostic prefix, including empty to clear the previous prefix.</param>
*)
METHOD INTERNAL FINAL Prepare
VAR_INPUT
	actual : SINT;
	testCase : ITestCase;
	message : WSTRING(255);
END_VAR
_Actual := actual;
_TestCase := testCase;
_Message := message;
END_METHOD

(*!
<summary>Reports the byte size of this concrete instance.</summary>
<description>
Includes inline fields and nested instances, but excludes separately allocated payloads.
Obtaining the size does not transfer ownership or validate an arbitrary address.
</description>
*)
{attribute 'monitoring' := 'call'}
PROPERTY SelfSize : ULINT
GET
SelfSize := XSIZEOF(THIS^);
END_GET
END_PROPERTY

(*!
<summary>Asserts equality with the expected value.</summary>
<description>
Records failure without interrupting the callback; preserves the message for the rest of the chain.
</description>
<param name="expected">Expected value converted by the compiler to SINT.</param>
*)
METHOD FINAL ToBe : REFERENCE TO SIntAssertionContext
VAR_INPUT
	expected : SINT;
END_VAR
IF _Actual <> expected THEN
	failComparison(
		expected := expected,
		expectation := "Expected: "
	);
END_IF

ToBe REF= THIS^;
END_METHOD

